screen "2#电梯状态画面" 800x600
   TextField "文本域_1" at 385,17 size 267x27; Text '-- 2#电梯状态总览'
   TextField "文本域_3" at 77,12 size 300x31; Text '电 梯 监 控 系 统'
   Button "按钮_7" at 555,516 size 117x66; TextOff '电梯状态总览'
      on Click: ActivateScreen("电梯状态总览画面", 0)
   Button "按钮_8" at 677,516 size 106x66; TextOff '退出系统'
      on Click: StopRuntime(0)
   Rectangle "矩形_237" at 73,319 size 44x21
      Appearance <- "输出_2号梯5层按钮指示灯"
   Rectangle "矩形_238" at 73,297 size 44x21
      Appearance <- "输出_2号梯6层按钮指示灯"
   Rectangle "矩形_239" at 73,275 size 44x21
      Appearance <- "输出_2号梯7层按钮指示灯"
   Rectangle "矩形_240" at 73,253 size 44x21
      Appearance <- "输出_2号梯8层按钮指示灯"
   Rectangle "矩形_241" at 73,231 size 44x21
      Appearance <- "输出_2号梯9层按钮指示灯"
   Rectangle "矩形_242" at 73,209 size 44x21
      Appearance <- "输出_2号梯10层按钮指示灯"
   Circle "圆_1" at 162,212 size 14x14
      Appearance <- "输出_10层下行呼梯按钮指示灯"
   Circle "圆_2" at 149,234 size 14x14
      Appearance <- "输出_9层上行呼梯按钮指示灯"
   Circle "圆_3" at 174,234 size 14x14
      Appearance <- "输出_9层下行呼梯按钮指示灯"
   Circle "圆_4" at 149,256 size 14x14
      Appearance <- "输出_8层上行呼梯按钮指示灯"
   Circle "圆_5" at 174,256 size 14x14
      Appearance <- "输出_8层下行呼梯按钮指示灯"
   Circle "圆_6" at 149,278 size 14x14
      Appearance <- "输出_7层上行呼梯按钮指示灯"
   Circle "圆_7" at 174,278 size 14x14
      Appearance <- "输出_7层下行呼梯按钮指示灯"
   Circle "圆_8" at 149,299 size 14x14
      Appearance <- "输出_6层上行呼梯按钮指示灯"
   Circle "圆_9" at 174,299 size 14x14
      Appearance <- "输出_6层下行呼梯按钮指示灯"
   Circle "圆_10" at 149,321 size 14x14
      Appearance <- "输出_5层上行呼梯按钮指示灯"
   Circle "圆_11" at 174,321 size 14x14
      Appearance <- "输出_5层下行呼梯按钮指示灯"
   Circle "圆_12" at 149,343 size 14x14
      Appearance <- "输出_4层上行呼梯按钮指示灯"
   Circle "圆_13" at 174,343 size 14x14
      Appearance <- "输出_4层下行呼梯按钮指示灯"
   Circle "圆_14" at 149,365 size 14x14
      Appearance <- "输出_3层上行呼梯按钮指示灯"
   Circle "圆_15" at 174,365 size 14x14
      Appearance <- "输出_3层下行呼梯按钮指示灯"
   Circle "圆_16" at 149,389 size 14x14
      Appearance <- "输出_2层上行呼梯按钮指示灯"
   Circle "圆_17" at 174,389 size 14x14
      Appearance <- "输出_2层下行呼梯按钮指示灯"
   Circle "圆_18" at 162,411 size 14x14
      Appearance <- "输出_1层上行呼梯按钮指示灯"
   TextField "文本域_41" at 75,440 size 45x23; Text '内呼'
   TextField "文本域_42" at 151,441 size 48x24; Text '外呼'
   Rectangle "矩形_233" at 73,407 size 44x21
      Appearance <- "输出_2号梯1层按钮指示灯"
   Rectangle "矩形_234" at 73,385 size 44x21
      Appearance <- "输出_2号梯2层按钮指示灯"
   Button "FB_Empty_Rectangular_1" at 80,409 size 29x18; TextOff 'Text'; PictureOff "FB_Empty_Rectangular_Released_256c"; PictureOn "FB_Empty_Rectangular_Pressed_256c"
      on Release: ResetBit("输入_2号梯轿内选层按钮1")
      on Press: SetBit("输入_2号梯轿内选层按钮1")
   Button "FB_Empty_Rectangular_2" at 81,387 size 29x18; TextOff 'Text'; PictureOff "FB_Empty_Rectangular_Released_256c"; PictureOn "FB_Empty_Rectangular_Pressed_256c"
      on Release: ResetBit("输入_2号梯轿内选层按钮2")
      on Press: SetBit("输入_2号梯轿内选层按钮2")
   Rectangle "矩形_235" at 73,363 size 44x21
      Appearance <- "输出_2号梯3层按钮指示灯"
   Button "FB_Empty_Rectangular_3" at 81,365 size 29x18; TextOff 'Text'; PictureOff "FB_Empty_Rectangular_Released_256c"; PictureOn "FB_Empty_Rectangular_Pressed_256c"
      on Release: ResetBit("输入_2号梯轿内选层按钮3")
      on Press: SetBit("输入_2号梯轿内选层按钮3")
   Rectangle "矩形_236" at 73,341 size 44x21
      Appearance <- "输出_2号梯4层按钮指示灯"
   Button "FB_Empty_Rectangular_4" at 81,343 size 29x18; TextOff 'Text'; PictureOff "FB_Empty_Rectangular_Released_256c"; PictureOn "FB_Empty_Rectangular_Pressed_256c"
      on Release: ResetBit("输入_2号梯轿内选层按钮4")
      on Press: SetBit("输入_2号梯轿内选层按钮4")
   Button "FB_Empty_Rectangular_5" at 81,321 size 29x18; TextOff 'Text'; PictureOff "FB_Empty_Rectangular_Released_256c"; PictureOn "FB_Empty_Rectangular_Pressed_256c"
      on Release: ResetBit("输入_2号梯轿内选层按钮5")
      on Press: SetBit("输入_2号梯轿内选层按钮5")
   Button "FB_Empty_Rectangular_6" at 81,299 size 29x18; TextOff 'Text'; PictureOff "FB_Empty_Rectangular_Released_256c"; PictureOn "FB_Empty_Rectangular_Pressed_256c"
      on Release: ResetBit("输入_2号梯轿内选层按钮6")
      on Press: SetBit("输入_2号梯轿内选层按钮6")
   Button "FB_Empty_Rectangular_7" at 81,277 size 29x18; TextOff 'Text'; PictureOff "FB_Empty_Rectangular_Released_256c"; PictureOn "FB_Empty_Rectangular_Pressed_256c"
      on Release: ResetBit("输入_2号梯轿内选层按钮7")
      on Press: SetBit("输入_2号梯轿内选层按钮7")
   Button "FB_Empty_Rectangular_8" at 81,255 size 29x18; TextOff 'Text'; PictureOff "FB_Empty_Rectangular_Released_256c"; PictureOn "FB_Empty_Rectangular_Pressed_256c"
      on Release: ResetBit("输入_2号梯轿内选层按钮8")
      on Press: SetBit("输入_2号梯轿内选层按钮8")
   Button "FB_Empty_Rectangular_9" at 81,233 size 29x18; TextOff 'Text'; PictureOff "FB_Empty_Rectangular_Released_256c"; PictureOn "FB_Empty_Rectangular_Pressed_256c"
      on Release: ResetBit("输入_2号梯轿内选层按钮9")
      on Press: SetBit("输入_2号梯轿内选层按钮9")
   Button "FB_Empty_Rectangular_10" at 81,211 size 29x18; TextOff 'Text'; PictureOff "FB_Empty_Rectangular_Released_256c"; PictureOn "FB_Empty_Rectangular_Pressed_256c"
      on Release: ResetBit("输入_2号梯轿内选层按钮10")
      on Press: SetBit("输入_2号梯轿内选层按钮10")
   TextField "文本域_14" at 88,409 size 14x19; Text '1'
   TextField "文本域_15" at 88,386 size 14x19; Text '2'
   TextField "文本域_16" at 88,363 size 14x19; Text '3'
   TextField "文本域_17" at 88,342 size 14x19; Text '4'
   TextField "文本域_18" at 88,320 size 14x19; Text '5'
   TextField "文本域_19" at 88,298 size 14x19; Text '6'
   TextField "文本域_20" at 88,276 size 14x19; Text '7'
   TextField "文本域_21" at 88,254 size 14x19; Text '8'
   TextField "文本域_22" at 88,232 size 14x19; Text '9'
   TextField "文本域_40" at 84,210 size 23x19; Text '10'
   Circle "圆_56" at 464,117 size 24x24
      Appearance <- "输出_2号梯满载指示"
   Circle "圆_57" at 574,117 size 24x24
      Appearance <- "输出_2号梯故障指示"
   Circle "圆_58" at 464,164 size 24x24
      Appearance <- "输出_2号梯照明指示"
   Circle "圆_59" at 349,120 size 24x24
      Appearance <- "输出_2号梯满载指示"
   Circle "圆_60" at 575,166 size 24x24
      Appearance <- "输出_2号梯风扇指示"
   TextField "文本域_47" at 383,122 size 37x19; Text '超重'
   TextField "文本域_48" at 498,120 size 61x23; Text '满载'
   TextField "文本域_49" at 608,118 size 50x28; Text '故障'
   TextField "文本域_50" at 502,167 size 54x26; Text '照明'
   TextField "文本域_51" at 609,162 size 58x28; Text '风扇'
   Circle "圆_73" at 215,119 size 24x24
      Appearance <- "输入_自动运行信号"
   TextField "文本域_68" at 246,120 size 87x20; Text '自动运行'
   Group "Group" at 310,468 size 40x20; PictureOn "FB_Left_Square_Pressed_256c"; PictureOff "FB_Left_Square_Released_256c"
   Group "Group_1" at 356,468 size 40x20; PictureOn "FB_Left_Square_Pressed_256c"; PictureOff "FB_Left_Square_Released_256c"
   TextField "文本域_69" at 245,167 size 127x20; Text '电梯准备就绪'
   Circle "圆_83" at 624,288 size 16x16
      Appearance <- "输出_2号梯开门继电器"
   Circle "圆_86" at 624,303 size 16x16
      Appearance <- "输出_2号梯关门继电器"
   Circle "圆_89" at 472,373 size 16x16
      Appearance <- "输入_2号梯开门到位"
   Circle "圆_92" at 472,389 size 16x16
      Appearance <- "输入_2号梯关门到位"
   Circle "圆_129" at 624,238 size 16x16
      Appearance <- "输出_2号梯电机启动信号"
   Circle "圆_132" at 624,253 size 16x16
      Appearance <- "输出_2号梯上行接触器"
   Circle "圆_135" at 624,268 size 16x16
      Appearance <- "输出_2号梯下行接触器"
   Circle "圆_19" at 215,163 size 24x24
      Appearance <- "输出_准备就绪信号"
   Circle "圆_95" at 624,358 size 16x16
      Appearance <- "输出_2号梯1级减速制动"
   Circle "圆_98" at 624,373 size 16x16
      Appearance <- "输出_2号梯2级减速制动"
   Circle "圆_101" at 624,388 size 16x16
      Appearance <- "输出_2号梯3级减速制动"
   Circle "圆_104" at 624,327 size 16x16
      Appearance <- "输出_2号梯低速接触器"
   Circle "圆_107" at 624,342 size 16x16
      Appearance <- "输出_2号梯高速接触器"
   Circle "圆_120" at 317,389 size 16x16
      Appearance <- "输入_2号梯轿厢门锁信号"
   Circle "圆_123" at 317,234 size 16x16
      Appearance <- "输入_2号梯10楼层门锁信号"
   Circle "圆_126" at 317,249 size 16x16
      Appearance <- "输入_2号梯9楼层门锁信号"
   Circle "圆_138" at 317,264 size 16x16
      Appearance <- "输入_2号梯8楼层门锁信号"
   Circle "圆_141" at 317,279 size 16x16
      Appearance <- "输入_2号梯7楼层门锁信号"
   Circle "圆_144" at 317,295 size 16x16
      Appearance <- "输入_2号梯6楼层门锁信号"
   Circle "圆_147" at 317,310 size 16x16
      Appearance <- "输入_2号梯5楼层门锁信号"
   Circle "圆_150" at 317,326 size 16x16
      Appearance <- "输入_2号梯4楼层门锁信号"
   Circle "圆_153" at 317,342 size 16x16
      Appearance <- "输入_2号梯3楼层门锁信号"
   Circle "圆_156" at 317,357 size 16x16
      Appearance <- "输入_2号梯2楼层门锁信号"
   Circle "圆_159" at 317,373 size 16x16
      Appearance <- "输入_2号梯1楼层门锁信号"
   Circle "圆_162" at 472,234 size 16x16
      Appearance <- "输入_2号梯上端站第2限位"
   Circle "圆_165" at 472,249 size 16x16
      Appearance <- "输入_2号梯上端站第1限位"
   Circle "圆_168" at 472,264 size 16x16
      Appearance <- "输入_2号梯上平层信号"
   Circle "圆_171" at 472,279 size 16x16
      Appearance <- "输入_2号梯下平层信号"
   Circle "圆_174" at 472,294 size 16x16
      Appearance <- "输入_2号梯下端站第2限位"
   Circle "圆_177" at 472,309 size 16x16
      Appearance <- "输入_2号梯下端站第1限位"
   Circle "圆_183" at 472,333 size 16x16
      Appearance <- "输入_2号梯检修信号"
   Circle "圆_186" at 472,348 size 16x16
      Appearance <- "输入_2号梯光幕信号"
   Rectangle "矩形_193" at 165,134 size 4x18
      Appearance <- "输出_2号梯LEDi"
   Rectangle "矩形_194" at 165,156 size 4x18
      Appearance <- "输出_2号梯LEDj"
   Rectangle "矩形_195" at 178,132 size 18x4
      Appearance <- "输出_2号梯LEDa"
   Rectangle "矩形_196" at 175,136 size 4x18
      Appearance <- "输出_2号梯LEDf"
   Rectangle "矩形_197" at 178,153 size 18x4
      Appearance <- "输出_2号梯LEDg"
   Rectangle "矩形_198" at 175,157 size 4x18
      Appearance <- "输出_2号梯LEDe"
   Rectangle "矩形_199" at 178,175 size 18x4
      Appearance <- "输出_2号梯LEDd"
   Rectangle "矩形_200" at 195,135 size 4x18
      Appearance <- "输出_2号梯LEDb"
   Rectangle "矩形_201" at 195,157 size 4x18
      Appearance <- "输出_2号梯LEDc"
   Rectangle "矩形_72" at 91,122 size 6x34
      Appearance <- "输出_2号梯上行指示"
   Polygon "多边形_5" at 79,118 size 15x17
      Appearance <- "输出_2号梯上行指示"
   Polygon "多边形_6" at 94,118 size 14x17
      Appearance <- "输出_2号梯上行指示"
   Rectangle "矩形_73" at 91,157 size 6x34
      Appearance <- "输出_2号梯下行指示"
   Polygon "多边形_1" at 77,179 size 17x15
      Appearance <- "输出_2号梯下行指示"
   Polygon "多边形_2" at 94,179 size 17x15
      Appearance <- "输出_2号梯下行指示"
   TextField "文本域_77" at 223,251 size 81x15; Text '9层门锁信号'
   TextField "文本域_78" at 223,266 size 81x15; Text '8层门锁信号'
   TextField "文本域_79" at 223,282 size 81x15; Text '7层门锁信号'
   TextField "文本域_80" at 223,298 size 81x15; Text '6层门锁信号'
   TextField "文本域_81" at 223,314 size 81x15; Text '5层门锁信号'
   TextField "文本域_83" at 223,329 size 81x15; Text '4层门锁信号'
   TextField "文本域_84" at 223,344 size 81x15; Text '3层门锁信号'
   TextField "文本域_85" at 223,360 size 81x15; Text '2层门锁信号'
   TextField "文本域_86" at 222,375 size 82x15; Text '1层门锁信号'
   TextField "文本域_87" at 223,391 size 81x15; Text '轿厢门锁信号'
   TextField "文本域_23" at 382,336 size 72x15; Text '检修开关'
   TextField "文本域_24" at 384,352 size 70x15; Text '光幕信号'
   TextField "文本域_82" at 351,237 size 103x15; Text '上端站第二限位'
   TextField "文本域_88" at 350,255 size 104x15; Text '上端站第一限位'
   TextField "文本域_89" at 372,270 size 82x15; Text '上平层信号'
   TextField "文本域_90" at 372,285 size 82x15; Text '下平层信号'
   TextField "文本域_91" at 350,299 size 104x15; Text '下端站第二限位'
   TextField "文本域_92" at 350,315 size 104x15; Text '下端站第一限位'
   TextField "文本域_13" at 362,372 size 93x15; Text '开门到位信号'
   TextField "文本域_25" at 362,388 size 93x15; Text '关门到位信号'
   TextField "文本域_97" at 525,289 size 92x15; Text '开门继电器'
   TextField "文本域_98" at 525,305 size 92x15; Text '关门继电器'
   TextField "文本域_104" at 525,270 size 92x15; Text '下行接触器'
   TextField "文本域_105" at 514,238 size 103x15; Text '电机启动信号'
   TextField "文本域_106" at 525,254 size 92x15; Text '上行接触器'
   TextField "文本域_99" at 504,374 size 114x15; Text '二级制动接触器'
   TextField "文本域_100" at 504,390 size 114x15; Text '三级制动接触器'
   TextField "文本域_101" at 504,357 size 114x15; Text '一级制动接触器'
   TextField "文本域_102" at 504,325 size 114x15; Text '低速运行接触器'
   TextField "文本域_103" at 504,341 size 114x15; Text '高速运行接触器'
   TextField "文本域_76" at 217,236 size 91x15; Text '10层门锁信号'
   Clock "时钟_1" at 664,57 size 101x57
   DateTimeField "日期/时间域_1" at 491,71 size 184x28
   TextField "文本域_26" at 278,421 size 142x19; Text '1号电梯开关门状态'
   Button "FB_Left_Square" at 310,468 size 20x20; TextOff 'Text'; PictureOff "FB_Left_Square_Released_256c"; PictureOn "FB_Left_Square_Pressed_256c"
      on Click: SetBit("输入_1号梯轿内开门按钮")
      Appearance <- "输入_2号梯轿内关门按钮"
   Button "FB_Right_Square" at 330,468 size 20x20; TextOff 'Text'; PictureOff "FB_Right_Square_Released_256c_2"; PictureOn "FB_Right_Square_Pressed_256c"
      on Click: SetBit("输入_1号梯轿内开门按钮")
      Appearance <- "输入_1号梯轿内开门按钮"
   Button "FB_Left_Square_1" at 376,468 size 20x20; TextOff 'Text'; PictureOff "FB_Left_Square_Released_256c"; PictureOn "FB_Left_Square_Pressed_256c"
      on Click: SetBit("输入_1号梯轿内关门按钮")
      Appearance <- "输入_2号梯轿内关门按钮"
   Button "FB_Right_Square_1" at 356,468 size 20x20; TextOff 'Text'; PictureOff "FB_Right_Square_Released_256c_2"; PictureOn "FB_Right_Square_Pressed_256c"
      on Click: SetBit("输入_1号梯轿内关门按钮")
      Appearance <- "输入_1号梯轿内关门按钮"

screen "3#电梯状态画面" 800x600
   TextField "文本域_1" at 385,17 size 263x27; Text '-- 3#电梯状态总览'
   TextField "文本域_3" at 82,12 size 295x31; Text '电 梯 监 控 系 统'
   Button "按钮_7" at 550,517 size 115x66; TextOff '电梯状态总览'
      on Click: ActivateScreen("电梯状态总览画面", 0)
   Button "按钮_8" at 671,517 size 106x66; TextOff '退出系统'
      on Click: StopRuntime(0)
   Group "Group" at 272,465 size 40x20; PictureOn "FB_Left_Square_Pressed_256c"; PictureOff "FB_Left_Square_Released_256c"
   Group "Group_1" at 324,465 size 40x20; PictureOn "FB_Left_Square_Pressed_256c"; PictureOff "FB_Left_Square_Released_256c"
   Rectangle "矩形_237" at 75,319 size 44x21
      Appearance <- "输出_3号梯5层按钮指示灯"
   Rectangle "矩形_238" at 75,297 size 44x21
      Appearance <- "输出_3号梯6层按钮指示灯"
   Rectangle "矩形_239" at 75,275 size 44x21
      Appearance <- "输出_3号梯7层按钮指示灯"
   Rectangle "矩形_240" at 75,253 size 44x21
      Appearance <- "输出_3号梯8层按钮指示灯"
   Rectangle "矩形_241" at 75,231 size 44x21
      Appearance <- "输出_3号梯9层按钮指示灯"
   Rectangle "矩形_242" at 75,209 size 44x21
      Appearance <- "输出_3号梯10层按钮指示灯"
   Circle "圆_1" at 164,212 size 14x14
      Appearance <- "输出_10层下行呼梯按钮指示灯"
   Circle "圆_2" at 151,232 size 14x14
      Appearance <- "输出_9层上行呼梯按钮指示灯"
   Circle "圆_3" at 176,232 size 14x14
      Appearance <- "输出_9层下行呼梯按钮指示灯"
   Circle "圆_4" at 151,254 size 14x14
      Appearance <- "输出_8层上行呼梯按钮指示灯"
   Circle "圆_5" at 176,254 size 14x14
      Appearance <- "输出_8层下行呼梯按钮指示灯"
   Circle "圆_6" at 151,277 size 14x14
      Appearance <- "输出_7层上行呼梯按钮指示灯"
   Circle "圆_7" at 176,277 size 14x14
      Appearance <- "输出_7层下行呼梯按钮指示灯"
   Circle "圆_8" at 151,299 size 14x14
      Appearance <- "输出_6层上行呼梯按钮指示灯"
   Circle "圆_9" at 176,299 size 14x14
      Appearance <- "输出_6层下行呼梯按钮指示灯"
   Circle "圆_10" at 151,322 size 14x14
      Appearance <- "输出_5层上行呼梯按钮指示灯"
   Circle "圆_11" at 176,322 size 14x14
      Appearance <- "输出_5层下行呼梯按钮指示灯"
   Circle "圆_12" at 151,345 size 14x14
      Appearance <- "输出_4层上行呼梯按钮指示灯"
   Circle "圆_13" at 176,345 size 14x14
      Appearance <- "输出_4层下行呼梯按钮指示灯"
   Circle "圆_14" at 151,367 size 14x14
      Appearance <- "输出_3层上行呼梯按钮指示灯"
   Circle "圆_15" at 176,367 size 14x14
      Appearance <- "输出_3层下行呼梯按钮指示灯"
   Circle "圆_16" at 151,389 size 14x14
      Appearance <- "输出_2层上行呼梯按钮指示灯"
   Circle "圆_17" at 176,389 size 14x14
      Appearance <- "输出_2层下行呼梯按钮指示灯"
   Circle "圆_18" at 163,411 size 14x14
      Appearance <- "输出_1层上行呼梯按钮指示灯"
   TextField "文本域_41" at 77,440 size 45x23; Text '内呼'
   TextField "文本域_42" at 152,440 size 45x23; Text '外呼'
   Rectangle "矩形_233" at 75,407 size 44x21
      Appearance <- "输出_3号梯1层按钮指示灯"
   Rectangle "矩形_234" at 75,385 size 44x21
      Appearance <- "输出_3号梯2层按钮指示灯"
   Button "FB_Empty_Rectangular_1" at 82,410 size 29x18; TextOff 'Text'; PictureOff "FB_Empty_Rectangular_Released_256c"; PictureOn "FB_Empty_Rectangular_Pressed_256c"
      on Release: ResetBit("输入_3号梯轿内选层按钮1")
      on Press: SetBit("输入_3号梯轿内选层按钮1")
      Appearance <- "输出_1号梯1层按钮指示灯"
   Button "FB_Empty_Rectangular_2" at 83,387 size 29x18; TextOff 'Text'; PictureOff "FB_Empty_Rectangular_Released_256c"; PictureOn "FB_Empty_Rectangular_Pressed_256c"
      on Release: ResetBit("输入_3号梯轿内选层按钮2")
      on Press: SetBit("输入_3号梯轿内选层按钮2")
   Rectangle "矩形_235" at 75,363 size 44x21
      Appearance <- "输出_3号梯3层按钮指示灯"
   Button "FB_Empty_Rectangular_3" at 83,365 size 29x18; TextOff 'Text'; PictureOff "FB_Empty_Rectangular_Released_256c"; PictureOn "FB_Empty_Rectangular_Pressed_256c"
      on Release: ResetBit("输入_3号梯轿内选层按钮3")
      on Press: SetBit("输入_3号梯轿内选层按钮3")
   Rectangle "矩形_236" at 75,341 size 44x21
      Appearance <- "输出_3号梯4层按钮指示灯"
   Button "FB_Empty_Rectangular_4" at 83,343 size 29x18; TextOff 'Text'; PictureOff "FB_Empty_Rectangular_Released_256c"; PictureOn "FB_Empty_Rectangular_Pressed_256c"
      on Release: ResetBit("输入_3号梯轿内选层按钮4")
      on Press: SetBit("输入_3号梯轿内选层按钮4")
   Button "FB_Empty_Rectangular_5" at 83,321 size 29x18; TextOff 'Text'; PictureOff "FB_Empty_Rectangular_Released_256c"; PictureOn "FB_Empty_Rectangular_Pressed_256c"
      on Release: ResetBit("输入_3号梯轿内选层按钮5")
      on Press: SetBit("输入_3号梯轿内选层按钮5")
   Button "FB_Empty_Rectangular_6" at 83,299 size 29x18; TextOff 'Text'; PictureOff "FB_Empty_Rectangular_Released_256c"; PictureOn "FB_Empty_Rectangular_Pressed_256c"
      on Release: ResetBit("输入_3号梯轿内选层按钮6")
      on Press: SetBit("输入_3号梯轿内选层按钮6")
   Button "FB_Empty_Rectangular_7" at 83,277 size 29x18; TextOff 'Text'; PictureOff "FB_Empty_Rectangular_Released_256c"; PictureOn "FB_Empty_Rectangular_Pressed_256c"
      on Release: ResetBit("输入_3号梯轿内选层按钮7")
      on Press: SetBit("输入_3号梯轿内选层按钮7")
   Button "FB_Empty_Rectangular_8" at 83,255 size 29x18; TextOff 'Text'; PictureOff "FB_Empty_Rectangular_Released_256c"; PictureOn "FB_Empty_Rectangular_Pressed_256c"
      on Release: ResetBit("输入_3号梯轿内选层按钮8")
      on Press: SetBit("输入_3号梯轿内选层按钮8")
   Button "FB_Empty_Rectangular_9" at 83,233 size 29x18; TextOff 'Text'; PictureOff "FB_Empty_Rectangular_Released_256c"; PictureOn "FB_Empty_Rectangular_Pressed_256c"
      on Release: ResetBit("输入_3号梯轿内选层按钮9")
      on Press: SetBit("输入_3号梯轿内选层按钮9")
   Button "FB_Empty_Rectangular_10" at 83,211 size 29x18; TextOff 'Text'; PictureOff "FB_Empty_Rectangular_Released_256c"; PictureOn "FB_Empty_Rectangular_Pressed_256c"
      on Release: ResetBit("输入_3号梯轿内选层按钮10")
      on Press: SetBit("输入_3号梯轿内选层按钮10")
   TextField "文本域_14" at 90,409 size 14x19; Text '1'
   TextField "文本域_15" at 90,386 size 14x19; Text '2'
   TextField "文本域_16" at 90,363 size 14x19; Text '3'
   TextField "文本域_17" at 90,342 size 14x19; Text '4'
   TextField "文本域_18" at 90,320 size 14x19; Text '5'
   TextField "文本域_19" at 90,298 size 14x19; Text '6'
   TextField "文本域_20" at 90,276 size 14x19; Text '7'
   TextField "文本域_21" at 90,254 size 14x19; Text '8'
   TextField "文本域_22" at 90,232 size 14x19; Text '9'
   TextField "文本域_40" at 86,210 size 23x19; Text '10'
   Circle "圆_56" at 476,117 size 24x24
      Appearance <- "输出_3号梯满载指示"
   Circle "圆_57" at 586,117 size 24x24
      Appearance <- "输出_3号梯故障指示"
   Circle "圆_58" at 476,166 size 24x24
      Appearance <- "输出_3号梯照明指示"
   Circle "圆_59" at 372,119 size 24x24
      Appearance <- "输出_3号梯满载指示"
   Circle "圆_60" at 587,168 size 24x24
      Appearance <- "输出_3号梯风扇指示"
   TextField "文本域_47" at 403,119 size 45x23; Text '超重'
   TextField "文本域_48" at 510,120 size 45x23; Text '满载'
   TextField "文本域_49" at 622,119 size 45x23; Text '故障'
   TextField "文本域_50" at 514,169 size 45x23; Text '照明'
   TextField "文本域_51" at 624,168 size 45x23; Text '风扇'
   Circle "圆_73" at 227,119 size 24x24
      Appearance <- "输入_自动运行信号"
   TextField "文本域_68" at 258,120 size 73x20; Text '自动运行'
   TextField "文本域_69" at 257,167 size 107x20; Text '电梯准备就绪'
   Circle "圆_83" at 625,280 size 16x16
      Appearance <- "输出_3号梯开门继电器"
   Circle "圆_86" at 625,295 size 16x16
      Appearance <- "输出_3号梯关门继电器"
   Circle "圆_89" at 477,363 size 16x16
      Appearance <- "输入_3号梯开门到位"
   Circle "圆_92" at 477,379 size 16x16
      Appearance <- "输入_3号梯关门到位"
   Circle "圆_129" at 624,229 size 16x16
      Appearance <- "输出_3号梯电机启动信号"
   Circle "圆_132" at 624,244 size 16x16
      Appearance <- "输出_3号梯上行接触器"
   Circle "圆_135" at 624,259 size 16x16
      Appearance <- "输出_3号梯下行接触器"
   Circle "圆_19" at 227,163 size 24x24
      Appearance <- "输出_准备就绪信号"
   Circle "圆_95" at 625,352 size 16x16
      Appearance <- "输出_3号梯1级减速制动"
   Circle "圆_98" at 625,367 size 16x16
      Appearance <- "输出_3号梯2级减速制动"
   Circle "圆_101" at 625,382 size 16x16
      Appearance <- "输出_3号梯3级减速制动"
   Circle "圆_104" at 625,321 size 16x16
      Appearance <- "输出_3号梯低速接触器"
   Circle "圆_107" at 625,336 size 16x16
      Appearance <- "输出_3号梯高速接触器"
   Circle "圆_120" at 324,378 size 16x16
      Appearance <- "输入_3号梯轿厢门锁信号"
   Circle "圆_123" at 324,228 size 16x16
      Appearance <- "输入_3号梯10楼层门锁信号"
   Circle "圆_126" at 324,243 size 16x16
      Appearance <- "输入_3号梯9楼层门锁信号"
   Circle "圆_138" at 324,258 size 16x16
      Appearance <- "输入_3号梯8楼层门锁信号"
   Circle "圆_141" at 324,273 size 16x16
      Appearance <- "输入_3号梯7楼层门锁信号"
   Circle "圆_144" at 324,288 size 16x16
      Appearance <- "输入_3号梯6楼层门锁信号"
   Circle "圆_147" at 324,303 size 16x16
      Appearance <- "输入_3号梯5楼层门锁信号"
   Circle "圆_150" at 324,318 size 16x16
      Appearance <- "输入_3号梯4楼层门锁信号"
   Circle "圆_153" at 324,333 size 16x16
      Appearance <- "输入_3号梯3楼层门锁信号"
   Circle "圆_156" at 324,348 size 16x16
      Appearance <- "输入_3号梯2楼层门锁信号"
   Circle "圆_159" at 324,363 size 16x16
      Appearance <- "输入_3号梯1楼层门锁信号"
   Circle "圆_162" at 476,228 size 16x16
      Appearance <- "输入_3号梯上端站第2限位"
   Circle "圆_165" at 476,243 size 16x16
      Appearance <- "输入_3号梯上端站第1限位"
   Circle "圆_168" at 476,258 size 16x16
      Appearance <- "输入_3号梯上平层信号"
   Circle "圆_171" at 476,273 size 16x16
      Appearance <- "输入_3号梯下平层信号"
   Circle "圆_174" at 476,288 size 16x16
      Appearance <- "输入_3号梯下端站第2限位"
   Circle "圆_177" at 476,303 size 16x16
      Appearance <- "输入_3号梯下端站第1限位"
   Circle "圆_183" at 476,327 size 16x16
      Appearance <- "输入_3号梯检修信号"
   Circle "圆_186" at 476,342 size 16x16
      Appearance <- "输入_3号梯光幕信号"
   Rectangle "矩形_193" at 167,134 size 4x18
      Appearance <- "输出_3号梯LEDi"
   Rectangle "矩形_194" at 167,156 size 4x18
      Appearance <- "输出_3号梯LEDj"
   Rectangle "矩形_195" at 180,132 size 18x4
      Appearance <- "输出_3号梯LEDa"
   Rectangle "矩形_196" at 177,136 size 4x18
      Appearance <- "输出_3号梯LEDf"
   Rectangle "矩形_197" at 180,153 size 18x4
      Appearance <- "输出_3号梯LEDg"
   Rectangle "矩形_198" at 177,157 size 4x18
      Appearance <- "输出_3号梯LEDe"
   Rectangle "矩形_199" at 180,175 size 18x4
      Appearance <- "输出_3号梯LEDd"
   Rectangle "矩形_200" at 197,135 size 4x18
      Appearance <- "输出_3号梯LEDb"
   Rectangle "矩形_201" at 197,157 size 4x18
      Appearance <- "输出_3号梯LEDc"
   Rectangle "矩形_72" at 93,122 size 6x34
      Appearance <- "输出_3号梯上行指示"
   Polygon "多边形_5" at 81,118 size 15x17
      Appearance <- "输出_3号梯上行指示"
   Polygon "多边形_6" at 96,118 size 14x17
      Appearance <- "输出_3号梯上行指示"
   Rectangle "矩形_73" at 93,157 size 6x34
      Appearance <- "输出_3号梯下行指示"
   Polygon "多边形_1" at 79,179 size 17x15
      Appearance <- "输出_3号梯下行指示"
   Polygon "多边形_2" at 96,179 size 17x15
      Appearance <- "输出_3号梯下行指示"
   TextField "文本域_23" at 388,326 size 72x15; Text '检修开关'
   TextField "文本域_24" at 390,342 size 70x15; Text '光幕信号'
   TextField "文本域_82" at 357,229 size 103x15; Text '上端站第二限位'
   TextField "文本域_88" at 356,245 size 104x15; Text '上端站第一限位'
   TextField "文本域_89" at 378,260 size 82x15; Text '上平层信号'
   TextField "文本域_90" at 378,275 size 82x15; Text '下平层信号'
   TextField "文本域_91" at 356,291 size 104x15; Text '下端站第二限位'
   TextField "文本域_92" at 356,307 size 104x15; Text '下端站第一限位'
   TextField "文本域_13" at 368,364 size 93x15; Text '开门到位信号'
   TextField "文本域_25" at 368,380 size 93x15; Text '关门到位信号'
   TextField "文本域_97" at 528,282 size 92x15; Text '开门继电器'
   TextField "文本域_98" at 528,298 size 92x15; Text '关门继电器'
   TextField "文本域_104" at 528,263 size 92x15; Text '下行接触器'
   TextField "文本域_105" at 517,231 size 103x15; Text '电机启动信号'
   TextField "文本域_106" at 528,247 size 92x15; Text '上行接触器'
   TextField "文本域_99" at 507,367 size 114x15; Text '二级制动接触器'
   TextField "文本域_100" at 507,383 size 114x15; Text '三级制动接触器'
   TextField "文本域_101" at 507,350 size 114x15; Text '一级制动接触器'
   TextField "文本域_102" at 507,318 size 114x15; Text '低速运行接触器'
   TextField "文本域_103" at 507,334 size 114x15; Text '高速运行接触器'
   TextField "文本域_76" at 219,229 size 91x15; Text '10层门锁信号'
   TextField "文本域_77" at 225,245 size 81x15; Text '9层门锁信号'
   TextField "文本域_78" at 225,260 size 81x15; Text '8层门锁信号'
   TextField "文本域_79" at 225,274 size 81x15; Text '7层门锁信号'
   TextField "文本域_80" at 225,289 size 81x15; Text '6层门锁信号'
   TextField "文本域_81" at 225,304 size 81x15; Text '5层门锁信号'
   TextField "文本域_83" at 225,319 size 81x15; Text '4层门锁信号'
   TextField "文本域_84" at 225,335 size 81x15; Text '3层门锁信号'
   TextField "文本域_85" at 225,350 size 81x15; Text '2层门锁信号'
   TextField "文本域_86" at 224,365 size 82x15; Text '1层门锁信号'
   TextField "文本域_87" at 225,380 size 81x15; Text '轿厢门锁信号'
   Clock "时钟_1" at 664,57 size 101x57
   DateTimeField "日期/时间域_1" at 491,71 size 184x28
   TextField "文本域_26" at 243,428 size 142x19; Text '1号电梯开关门状态'
   Button "FB_Left_Square" at 272,465 size 20x20; TextOff 'Text'; PictureOff "FB_Left_Square_Released_256c"; PictureOn "FB_Left_Square_Pressed_256c"
      on Click: SetBit("输入_1号梯轿内开门按钮")
      Appearance <- "输入_3号梯轿内开门按钮"
   Button "FB_Right_Square" at 292,465 size 20x20; TextOff 'Text'; PictureOff "FB_Right_Square_Released_256c_3"; PictureOn "FB_Right_Square_Pressed_256c"
      on Click: SetBit("输入_1号梯轿内开门按钮")
      Appearance <- "输入_1号梯轿内开门按钮"
   Button "FB_Left_Square_1" at 344,465 size 20x20; TextOff 'Text'; PictureOff "FB_Left_Square_Released_256c"; PictureOn "FB_Left_Square_Pressed_256c"
      on Click: SetBit("输入_1号梯轿内关门按钮")
      Appearance <- "输入_3号梯轿内关门按钮"
   Button "FB_Right_Square_1" at 324,465 size 20x20; TextOff 'Text'; PictureOff "FB_Right_Square_Released_256c_3"; PictureOn "FB_Right_Square_Pressed_256c"
      on Click: SetBit("输入_1号梯轿内关门按钮")
      Appearance <- "输入_1号梯轿内关门按钮"

screen "4#电梯状态画面" 800x600
   TextField "文本域_1" at 385,17 size 287x27; Text '-- 4#电梯状态总览'
   TextField "文本域_3" at 71,12 size 306x31; Text '电 梯 监 控 系 统'
   Button "按钮_7" at 538,519 size 118x66; TextOff '电梯状态总览'
      on Click: ActivateScreen("电梯状态总览画面", 0)
   Button "按钮_8" at 664,519 size 106x66; TextOff '退出系统'
      on Click: StopRuntime(0)
   Group "Group" at 303,439 size 40x20; PictureOn "FB_Left_Square_Pressed_256c"; PictureOff "FB_Left_Square_Released_256c"
   Group "Group_1" at 349,439 size 40x20; PictureOn "FB_Left_Square_Pressed_256c"; PictureOff "FB_Left_Square_Released_256c"
   Rectangle "矩形_237" at 75,315 size 44x21
      Appearance <- "输出_4号梯5层按钮指示灯"
   Rectangle "矩形_238" at 75,293 size 44x21
      Appearance <- "输出_4号梯6层按钮指示灯"
   Rectangle "矩形_239" at 75,271 size 44x21
      Appearance <- "输出_4号梯7层按钮指示灯"
   Rectangle "矩形_240" at 75,249 size 44x21
      Appearance <- "输出_4号梯8层按钮指示灯"
   Rectangle "矩形_241" at 75,227 size 44x21
      Appearance <- "输出_4号梯9层按钮指示灯"
   Rectangle "矩形_242" at 75,205 size 44x21
      Appearance <- "输出_4号梯10层按钮指示灯"
   Circle "圆_1" at 162,208 size 14x14
      Appearance <- "输出_10层下行呼梯按钮指示灯"
   Circle "圆_2" at 151,230 size 14x14
      Appearance <- "输出_9层上行呼梯按钮指示灯"
   Circle "圆_3" at 176,230 size 14x14
      Appearance <- "输出_9层下行呼梯按钮指示灯"
   Circle "圆_4" at 151,251 size 14x14
      Appearance <- "输出_8层上行呼梯按钮指示灯"
   Circle "圆_5" at 176,251 size 14x14
      Appearance <- "输出_8层下行呼梯按钮指示灯"
   Circle "圆_6" at 151,273 size 14x14
      Appearance <- "输出_7层上行呼梯按钮指示灯"
   Circle "圆_7" at 176,273 size 14x14
      Appearance <- "输出_7层下行呼梯按钮指示灯"
   Circle "圆_8" at 151,296 size 14x14
      Appearance <- "输出_6层上行呼梯按钮指示灯"
   Circle "圆_9" at 176,296 size 14x14
      Appearance <- "输出_6层下行呼梯按钮指示灯"
   Circle "圆_10" at 151,318 size 14x14
      Appearance <- "输出_5层上行呼梯按钮指示灯"
   Circle "圆_11" at 176,318 size 14x14
      Appearance <- "输出_5层下行呼梯按钮指示灯"
   Circle "圆_12" at 151,341 size 14x14
      Appearance <- "输出_4层上行呼梯按钮指示灯"
   Circle "圆_13" at 176,341 size 14x14
      Appearance <- "输出_4层下行呼梯按钮指示灯"
   Circle "圆_14" at 151,364 size 14x14
      Appearance <- "输出_3层上行呼梯按钮指示灯"
   Circle "圆_15" at 176,364 size 14x14
      Appearance <- "输出_3层下行呼梯按钮指示灯"
   Circle "圆_16" at 151,385 size 14x14
      Appearance <- "输出_2层上行呼梯按钮指示灯"
   Circle "圆_17" at 176,385 size 14x14
      Appearance <- "输出_2层下行呼梯按钮指示灯"
   Circle "圆_18" at 164,407 size 14x14
      Appearance <- "输出_1层上行呼梯按钮指示灯"
   TextField "文本域_41" at 77,436 size 45x23; Text '内呼'
   TextField "文本域_42" at 145,434 size 45x23; Text '外呼'
   Rectangle "矩形_233" at 75,403 size 44x21
      Appearance <- "输出_4号梯1层按钮指示灯"
   Rectangle "矩形_234" at 75,381 size 44x21
      Appearance <- "输出_4号梯2层按钮指示灯"
   Button "FB_Empty_Rectangular_1" at 82,406 size 29x18; TextOff 'Text'; PictureOff "FB_Empty_Rectangular_Released_256c"; PictureOn "FB_Empty_Rectangular_Pressed_256c"
      on Release: ResetBit("输入_1号梯轿内选层按钮1")
      on Press: SetBit("输入_1号梯轿内选层按钮1")
   Button "FB_Empty_Rectangular_2" at 83,383 size 29x18; TextOff 'Text'; PictureOff "FB_Empty_Rectangular_Released_256c"; PictureOn "FB_Empty_Rectangular_Pressed_256c"
      on Release: ResetBit("输入_1号梯轿内选层按钮2")
      on Press: SetBit("输入_1号梯轿内选层按钮2")
   Rectangle "矩形_235" at 75,359 size 44x21
      Appearance <- "输出_4号梯3层按钮指示灯"
   Button "FB_Empty_Rectangular_3" at 83,361 size 29x18; TextOff 'Text'; PictureOff "FB_Empty_Rectangular_Released_256c"; PictureOn "FB_Empty_Rectangular_Pressed_256c"
      on Release: ResetBit("输入_1号梯轿内选层按钮3")
      on Press: SetBit("输入_1号梯轿内选层按钮3")
   Rectangle "矩形_236" at 75,337 size 44x21
      Appearance <- "输出_4号梯4层按钮指示灯"
   Button "FB_Empty_Rectangular_4" at 83,339 size 29x18; TextOff 'Text'; PictureOff "FB_Empty_Rectangular_Released_256c"; PictureOn "FB_Empty_Rectangular_Pressed_256c"
      on Release: ResetBit("输入_1号梯轿内选层按钮4")
      on Press: SetBit("输入_1号梯轿内选层按钮4")
   Button "FB_Empty_Rectangular_5" at 83,317 size 29x18; TextOff 'Text'; PictureOff "FB_Empty_Rectangular_Released_256c"; PictureOn "FB_Empty_Rectangular_Pressed_256c"
      on Release: ResetBit("输入_1号梯轿内选层按钮5")
      on Press: SetBit("输入_1号梯轿内选层按钮5")
   Button "FB_Empty_Rectangular_6" at 83,295 size 29x18; TextOff 'Text'; PictureOff "FB_Empty_Rectangular_Released_256c"; PictureOn "FB_Empty_Rectangular_Pressed_256c"
      on Release: ResetBit("输入_1号梯轿内选层按钮6")
      on Press: SetBit("输入_1号梯轿内选层按钮6")
   Button "FB_Empty_Rectangular_7" at 83,273 size 29x18; TextOff 'Text'; PictureOff "FB_Empty_Rectangular_Released_256c"; PictureOn "FB_Empty_Rectangular_Pressed_256c"
      on Release: ResetBit("输入_1号梯轿内选层按钮7")
      on Press: SetBit("输入_1号梯轿内选层按钮7")
   Button "FB_Empty_Rectangular_8" at 83,251 size 29x18; TextOff 'Text'; PictureOff "FB_Empty_Rectangular_Released_256c"; PictureOn "FB_Empty_Rectangular_Pressed_256c"
      on Release: ResetBit("输入_1号梯轿内选层按钮8")
      on Press: SetBit("输入_1号梯轿内选层按钮8")
   Button "FB_Empty_Rectangular_9" at 83,229 size 29x18; TextOff 'Text'; PictureOff "FB_Empty_Rectangular_Released_256c"; PictureOn "FB_Empty_Rectangular_Pressed_256c"
      on Release: ResetBit("输入_1号梯轿内选层按钮9")
      on Press: SetBit("输入_1号梯轿内选层按钮9")
   Button "FB_Empty_Rectangular_10" at 83,207 size 29x18; TextOff 'Text'; PictureOff "FB_Empty_Rectangular_Released_256c"; PictureOn "FB_Empty_Rectangular_Pressed_256c"
      on Release: ResetBit("输入_1号梯轿内选层按钮10")
      on Press: SetBit("输入_1号梯轿内选层按钮10")
   TextField "文本域_14" at 90,405 size 14x19; Text '1'
   TextField "文本域_15" at 90,382 size 14x19; Text '2'
   TextField "文本域_16" at 90,359 size 14x19; Text '3'
   TextField "文本域_17" at 90,338 size 14x19; Text '4'
   TextField "文本域_18" at 90,316 size 14x19; Text '5'
   TextField "文本域_19" at 90,294 size 14x19; Text '6'
   TextField "文本域_20" at 90,272 size 14x19; Text '7'
   TextField "文本域_21" at 90,250 size 14x19; Text '8'
   TextField "文本域_22" at 90,228 size 14x19; Text '9'
   TextField "文本域_40" at 86,206 size 23x19; Text '10'
   Circle "圆_56" at 470,112 size 24x24
      Appearance <- "输出_4号梯满载指示"
   Circle "圆_57" at 580,112 size 24x24
      Appearance <- "输出_4号梯故障指示"
   Circle "圆_58" at 470,156 size 24x24
      Appearance <- "输出_4号梯照明指示"
   Circle "圆_59" at 368,114 size 24x24
      Appearance <- "输出_4号梯满载指示"
   Circle "圆_60" at 581,158 size 24x24
      Appearance <- "输出_4号梯风扇指示"
   TextField "文本域_47" at 397,114 size 45x23; Text '超重'
   TextField "文本域_48" at 504,115 size 45x23; Text '满载'
   TextField "文本域_49" at 616,114 size 45x23; Text '故障'
   TextField "文本域_50" at 508,159 size 45x23; Text '照明'
   TextField "文本域_51" at 618,159 size 45x23; Text '风扇'
   Circle "圆_73" at 221,114 size 24x24
      Appearance <- "输入_自动运行信号"
   TextField "文本域_68" at 252,115 size 73x20; Text '自动运行'
   TextField "文本域_69" at 254,162 size 107x20; Text '电梯准备就绪'
   Circle "圆_83" at 476,348 size 16x16
      Appearance <- "输出_4号梯开门继电器"
   Circle "圆_86" at 476,363 size 16x16
      Appearance <- "输出_4号梯关门继电器"
   Circle "圆_89" at 626,267 size 16x16
      Appearance <- "输入_4号梯开门到位"
   Circle "圆_92" at 626,283 size 16x16
      Appearance <- "输入_4号梯关门到位"
   Circle "圆_129" at 626,214 size 16x16
      Appearance <- "输出_4号梯电机启动信号"
   Circle "圆_132" at 626,229 size 16x16
      Appearance <- "输出_4号梯上行接触器"
   Circle "圆_135" at 626,244 size 16x16
      Appearance <- "输出_4号梯下行接触器"
   Circle "圆_19" at 221,158 size 24x24
      Appearance <- "输出_准备就绪信号"
   Circle "圆_95" at 627,338 size 16x16
      Appearance <- "输出_4号梯1级减速制动"
   Circle "圆_98" at 627,353 size 16x16
      Appearance <- "输出_4号梯2级减速制动"
   Circle "圆_101" at 627,368 size 16x16
      Appearance <- "输出_4号梯3级减速制动"
   Circle "圆_104" at 627,307 size 16x16
      Appearance <- "输出_4号梯低速接触器"
   Circle "圆_107" at 627,322 size 16x16
      Appearance <- "输出_4号梯高速接触器"
   Circle "圆_120" at 331,366 size 16x16
      Appearance <- "输入_4号梯轿厢门锁信号"
   Circle "圆_123" at 331,214 size 16x16
      Appearance <- "输入_4号梯10楼层门锁信号"
   Circle "圆_126" at 331,229 size 16x16
      Appearance <- "输入_4号梯9楼层门锁信号"
   Circle "圆_138" at 331,244 size 16x16
      Appearance <- "输入_4号梯8楼层门锁信号"
   Circle "圆_141" at 331,259 size 16x16
      Appearance <- "输入_4号梯7楼层门锁信号"
   Circle "圆_144" at 331,274 size 16x16
      Appearance <- "输入_4号梯6楼层门锁信号"
   Circle "圆_147" at 331,289 size 16x16
      Appearance <- "输入_4号梯5楼层门锁信号"
   Circle "圆_150" at 331,304 size 16x16
      Appearance <- "输入_4号梯4楼层门锁信号"
   Circle "圆_153" at 331,319 size 16x16
      Appearance <- "输入_4号梯3楼层门锁信号"
   Circle "圆_156" at 331,334 size 16x16
      Appearance <- "输入_4号梯2楼层门锁信号"
   Circle "圆_159" at 331,350 size 16x16
      Appearance <- "输入_4号梯1楼层门锁信号"
   Circle "圆_162" at 476,212 size 16x16
      Appearance <- "输入_4号梯上端站第2限位"
   Circle "圆_165" at 476,227 size 16x16
      Appearance <- "输入_4号梯上端站第1限位"
   Circle "圆_168" at 476,242 size 16x16
      Appearance <- "输入_4号梯上平层信号"
   Circle "圆_171" at 476,257 size 16x16
      Appearance <- "输入_4号梯下平层信号"
   Circle "圆_174" at 476,272 size 16x16
      Appearance <- "输入_4号梯下端站第2限位"
   Circle "圆_177" at 476,287 size 16x16
      Appearance <- "输入_4号梯下端站第1限位"
   Circle "圆_183" at 476,312 size 16x16
      Appearance <- "输入_4号梯检修信号"
   Circle "圆_186" at 476,327 size 16x16
      Appearance <- "输入_4号梯光幕信号"
   Rectangle "矩形_193" at 167,130 size 4x18
      Appearance <- "输出_4号梯LEDi"
   Rectangle "矩形_194" at 167,152 size 4x18
      Appearance <- "输出_4号梯LEDj"
   Rectangle "矩形_195" at 180,128 size 18x4
      Appearance <- "输出_4号梯LEDa"
   Rectangle "矩形_196" at 177,132 size 4x18
      Appearance <- "输出_4号梯LEDf"
   Rectangle "矩形_197" at 180,149 size 18x4
      Appearance <- "输出_4号梯LEDg"
   Rectangle "矩形_198" at 177,153 size 4x18
      Appearance <- "输出_4号梯LEDe"
   Rectangle "矩形_199" at 180,171 size 18x4
      Appearance <- "输出_4号梯LEDd"
   Rectangle "矩形_200" at 197,131 size 4x18
      Appearance <- "输出_4号梯LEDb"
   Rectangle "矩形_201" at 197,153 size 4x18
      Appearance <- "输出_4号梯LEDc"
   Rectangle "矩形_72" at 93,118 size 6x34
      Appearance <- "输出_4号梯上行指示"
   Polygon "多边形_5" at 81,114 size 15x17
      Appearance <- "输出_4号梯上行指示"
   Polygon "多边形_6" at 96,114 size 14x17
      Appearance <- "输出_4号梯上行指示"
   Rectangle "矩形_73" at 93,153 size 6x34
      Appearance <- "输出_4号梯下行指示"
   Polygon "多边形_1" at 79,175 size 17x15
      Appearance <- "输出_4号梯下行指示"
   Polygon "多边形_2" at 96,175 size 17x15
      Appearance <- "输出_4号梯下行指示"
   TextField "文本域_77" at 225,231 size 81x15; Text '9层门锁信号'
   TextField "文本域_78" at 225,245 size 81x15; Text '8层门锁信号'
   TextField "文本域_79" at 225,260 size 81x15; Text '7层门锁信号'
   TextField "文本域_80" at 225,275 size 81x15; Text '6层门锁信号'
   TextField "文本域_81" at 225,290 size 81x15; Text '5层门锁信号'
   TextField "文本域_83" at 225,306 size 81x15; Text '4层门锁信号'
   TextField "文本域_84" at 225,322 size 81x15; Text '3层门锁信号'
   TextField "文本域_85" at 225,337 size 81x15; Text '2层门锁信号'
   TextField "文本域_86" at 224,354 size 82x15; Text '1层门锁信号'
   TextField "文本域_87" at 220,369 size 86x15; Text '轿厢门锁信号'
   TextField "文本域_23" at 399,312 size 72x15; Text '检修开关'
   TextField "文本域_24" at 401,328 size 70x15; Text '光幕信号'
   TextField "文本域_82" at 368,215 size 103x15; Text '上端站第二限位'
   TextField "文本域_88" at 367,231 size 104x15; Text '上端站第一限位'
   TextField "文本域_89" at 389,246 size 82x15; Text '上平层信号'
   TextField "文本域_90" at 389,261 size 82x15; Text '下平层信号'
   TextField "文本域_91" at 367,275 size 104x15; Text '下端站第二限位'
   TextField "文本域_92" at 367,291 size 104x15; Text '下端站第一限位'
   TextField "文本域_13" at 379,348 size 93x15; Text '开门到位信号'
   TextField "文本域_25" at 379,364 size 93x15; Text '关门到位信号'
   TextField "文本域_97" at 531,267 size 92x15; Text '开门继电器'
   TextField "文本域_98" at 531,283 size 92x15; Text '关门继电器'
   TextField "文本域_104" at 531,248 size 92x15; Text '下行接触器'
   TextField "文本域_105" at 520,216 size 103x15; Text '电机启动信号'
   TextField "文本域_106" at 531,232 size 92x15; Text '上行接触器'
   TextField "文本域_99" at 510,352 size 114x15; Text '二级制动接触器'
   TextField "文本域_100" at 510,368 size 114x15; Text '三级制动接触器'
   TextField "文本域_101" at 510,335 size 114x15; Text '一级制动接触器'
   TextField "文本域_102" at 510,303 size 114x15; Text '低速运行接触器'
   TextField "文本域_103" at 510,319 size 114x15; Text '高速运行接触器'
   TextField "文本域_76" at 219,214 size 91x15; Text '10层门锁信号'
   Clock "时钟_1" at 664,57 size 101x57
   DateTimeField "日期/时间域_1" at 491,71 size 184x28
   TextField "文本域_26" at 269,403 size 142x19; Text '1号电梯开关门状态'
   Button "FB_Left_Square" at 303,439 size 20x20; TextOff 'Text'; PictureOff "FB_Left_Square_Released_256c"; PictureOn "FB_Left_Square_Pressed_256c"
      on Click: SetBit("输入_1号梯轿内开门按钮")
      Appearance <- "输入_4号梯轿内开门按钮"
   Button "FB_Right_Square" at 323,439 size 20x20; TextOff 'Text'; PictureOff "FB_Right_Square_Released_256c_4"; PictureOn "FB_Right_Square_Pressed_256c"
      on Click: SetBit("输入_1号梯轿内开门按钮")
      Appearance <- "输入_1号梯轿内开门按钮"
   Button "FB_Left_Square_1" at 369,439 size 20x20; TextOff 'Text'; PictureOff "FB_Left_Square_Released_256c"; PictureOn "FB_Left_Square_Pressed_256c"
      on Click: SetBit("输入_1号梯轿内关门按钮")
      Appearance <- "输入_4号梯轿内关门按钮"
   Button "FB_Right_Square_1" at 349,439 size 20x20; TextOff 'Text'; PictureOff "FB_Right_Square_Released_256c_4"; PictureOn "FB_Right_Square_Pressed_256c"
      on Click: SetBit("输入_1号梯轿内关门按钮")
      Appearance <- "输入_1号梯轿内关门按钮"

screen "5#电梯状态画面" 800x600
   TextField "文本域_1" at 385,17 size 274x27; Text '-- 5#电梯状态总览'
   TextField "文本域_3" at 76,12 size 301x31; Text '电 梯 监 控 系 统'
   Button "按钮_7" at 547,518 size 121x66; TextOff '电梯状态总览'
      on Click: ActivateScreen("电梯状态总览画面", 0)
   Button "按钮_8" at 675,518 size 106x66; TextOff '退出系统'
      on Click: StopRuntime(0)
   Group "Group" at 284,442 size 40x20; PictureOn "FB_Left_Square_Pressed_256c"; PictureOff "FB_Left_Square_Released_256c"
   Group "Group_1" at 330,442 size 40x20; PictureOn "FB_Left_Square_Pressed_256c"; PictureOff "FB_Left_Square_Released_256c"
   Rectangle "矩形_237" at 75,319 size 44x21
      Appearance <- "输出_5号梯5层按钮指示灯"
   Rectangle "矩形_238" at 75,297 size 44x21
      Appearance <- "输出_5号梯6层按钮指示灯"
   Rectangle "矩形_239" at 75,275 size 44x21
      Appearance <- "输出_5号梯7层按钮指示灯"
   Rectangle "矩形_240" at 75,253 size 44x21
      Appearance <- "输出_5号梯8层按钮指示灯"
   Rectangle "矩形_241" at 75,231 size 44x21
      Appearance <- "输出_5号梯9层按钮指示灯"
   Rectangle "矩形_242" at 75,209 size 44x21
      Appearance <- "输出_5号梯10层按钮指示灯"
   Circle "圆_1" at 163,212 size 14x14
      Appearance <- "输出_10层下行呼梯按钮指示灯"
   Circle "圆_2" at 151,233 size 14x14
      Appearance <- "输出_9层上行呼梯按钮指示灯"
   Circle "圆_3" at 176,233 size 14x14
      Appearance <- "输出_9层下行呼梯按钮指示灯"
   Circle "圆_4" at 151,254 size 14x14
      Appearance <- "输出_8层上行呼梯按钮指示灯"
   Circle "圆_5" at 176,254 size 14x14
      Appearance <- "输出_8层下行呼梯按钮指示灯"
   Circle "圆_6" at 151,277 size 14x14
      Appearance <- "输出_7层上行呼梯按钮指示灯"
   Circle "圆_7" at 176,277 size 14x14
      Appearance <- "输出_7层下行呼梯按钮指示灯"
   Circle "圆_8" at 151,299 size 14x14
      Appearance <- "输出_6层上行呼梯按钮指示灯"
   Circle "圆_9" at 176,299 size 14x14
      Appearance <- "输出_6层下行呼梯按钮指示灯"
   Circle "圆_10" at 151,322 size 14x14
      Appearance <- "输出_5层上行呼梯按钮指示灯"
   Circle "圆_11" at 176,322 size 14x14
      Appearance <- "输出_5层下行呼梯按钮指示灯"
   Circle "圆_12" at 151,345 size 14x14
      Appearance <- "输出_4层上行呼梯按钮指示灯"
   Circle "圆_13" at 176,345 size 14x14
      Appearance <- "输出_4层下行呼梯按钮指示灯"
   Circle "圆_14" at 151,366 size 14x14
      Appearance <- "输出_3层上行呼梯按钮指示灯"
   Circle "圆_15" at 176,366 size 14x14
      Appearance <- "输出_3层下行呼梯按钮指示灯"
   Circle "圆_16" at 151,389 size 14x14
      Appearance <- "输出_2层上行呼梯按钮指示灯"
   Circle "圆_17" at 176,389 size 14x14
      Appearance <- "输出_2层下行呼梯按钮指示灯"
   Circle "圆_18" at 163,411 size 14x14
      Appearance <- "输出_1层上行呼梯按钮指示灯"
   TextField "文本域_41" at 77,440 size 45x23; Text '内呼'
   TextField "文本域_42" at 153,438 size 45x23; Text '外呼'
   Rectangle "矩形_233" at 75,407 size 44x21
      Appearance <- "输出_5号梯1层按钮指示灯"
   Rectangle "矩形_234" at 75,385 size 44x21
      Appearance <- "输出_5号梯2层按钮指示灯"
   Button "FB_Empty_Rectangular_1" at 82,410 size 29x18; TextOff 'Text'; PictureOff "FB_Empty_Rectangular_Released_256c"; PictureOn "FB_Empty_Rectangular_Pressed_256c"
      on Release: ResetBit("输入_5号梯轿内选层按钮1")
      on Press: SetBit("输入_5号梯轿内选层按钮1")
   Button "FB_Empty_Rectangular_2" at 83,387 size 29x18; TextOff 'Text'; PictureOff "FB_Empty_Rectangular_Released_256c"; PictureOn "FB_Empty_Rectangular_Pressed_256c"
      on Release: ResetBit("输入_5号梯轿内选层按钮2")
      on Press: SetBit("输入_5号梯轿内选层按钮2")
   Rectangle "矩形_235" at 75,363 size 44x21
      Appearance <- "输出_5号梯3层按钮指示灯"
   Button "FB_Empty_Rectangular_3" at 83,365 size 29x18; TextOff 'Text'; PictureOff "FB_Empty_Rectangular_Released_256c"; PictureOn "FB_Empty_Rectangular_Pressed_256c"
      on Release: ResetBit("输入_5号梯轿内选层按钮3")
      on Press: SetBit("输入_5号梯轿内选层按钮3")
   Rectangle "矩形_236" at 75,341 size 44x21
      Appearance <- "输出_5号梯4层按钮指示灯"
   Button "FB_Empty_Rectangular_4" at 83,343 size 29x18; TextOff 'Text'; PictureOff "FB_Empty_Rectangular_Released_256c"; PictureOn "FB_Empty_Rectangular_Pressed_256c"
      on Release: ResetBit("输入_5号梯轿内选层按钮4")
      on Press: SetBit("输入_5号梯轿内选层按钮4")
   Button "FB_Empty_Rectangular_5" at 83,321 size 29x18; TextOff 'Text'; PictureOff "FB_Empty_Rectangular_Released_256c"; PictureOn "FB_Empty_Rectangular_Pressed_256c"
      on Release: ResetBit("输入_5号梯轿内选层按钮5")
      on Press: SetBit("输入_5号梯轿内选层按钮5")
   Button "FB_Empty_Rectangular_6" at 83,299 size 29x18; TextOff 'Text'; PictureOff "FB_Empty_Rectangular_Released_256c"; PictureOn "FB_Empty_Rectangular_Pressed_256c"
      on Release: ResetBit("输入_5号梯轿内选层按钮6")
      on Press: SetBit("输入_5号梯轿内选层按钮6")
   Button "FB_Empty_Rectangular_7" at 83,277 size 29x18; TextOff 'Text'; PictureOff "FB_Empty_Rectangular_Released_256c"; PictureOn "FB_Empty_Rectangular_Pressed_256c"
      on Release: ResetBit("输入_5号梯轿内选层按钮7")
      on Press: SetBit("输入_5号梯轿内选层按钮7")
   Button "FB_Empty_Rectangular_8" at 83,255 size 29x18; TextOff 'Text'; PictureOff "FB_Empty_Rectangular_Released_256c"; PictureOn "FB_Empty_Rectangular_Pressed_256c"
      on Release: ResetBit("输入_5号梯轿内选层按钮8")
      on Press: SetBit("输入_5号梯轿内选层按钮8")
   Button "FB_Empty_Rectangular_9" at 83,233 size 29x18; TextOff 'Text'; PictureOff "FB_Empty_Rectangular_Released_256c"; PictureOn "FB_Empty_Rectangular_Pressed_256c"
      on Release: ResetBit("输入_5号梯轿内选层按钮9")
      on Press: SetBit("输入_5号梯轿内选层按钮9")
   Button "FB_Empty_Rectangular_10" at 83,211 size 29x18; TextOff 'Text'; PictureOff "FB_Empty_Rectangular_Released_256c"; PictureOn "FB_Empty_Rectangular_Pressed_256c"
      on Release: ResetBit("输入_5号梯轿内选层按钮10")
      on Press: SetBit("输入_5号梯轿内选层按钮10")
   TextField "文本域_14" at 90,409 size 14x19; Text '1'
   TextField "文本域_15" at 90,386 size 14x19; Text '2'
   TextField "文本域_16" at 90,363 size 14x19; Text '3'
   TextField "文本域_17" at 90,342 size 14x19; Text '4'
   TextField "文本域_18" at 90,320 size 14x19; Text '5'
   TextField "文本域_19" at 90,298 size 14x19; Text '6'
   TextField "文本域_20" at 90,276 size 14x19; Text '7'
   TextField "文本域_21" at 90,254 size 14x19; Text '8'
   TextField "文本域_22" at 90,232 size 14x19; Text '9'
   TextField "文本域_40" at 86,210 size 23x19; Text '10'
   Circle "圆_56" at 475,117 size 24x24
      Appearance <- "输出_5号梯满载指示"
   Circle "圆_57" at 585,117 size 24x24
      Appearance <- "输出_5号梯故障指示"
   Circle "圆_58" at 473,163 size 24x24
      Appearance <- "输出_5号梯照明指示"
   Circle "圆_59" at 368,122 size 24x24
      Appearance <- "输出_5号梯满载指示"
   Circle "圆_60" at 584,165 size 24x24
      Appearance <- "输出_5号梯风扇指示"
   TextField "文本域_47" at 402,119 size 45x23; Text '超重'
   TextField "文本域_48" at 509,120 size 45x23; Text '满载'
   TextField "文本域_49" at 621,119 size 45x23; Text '故障'
   TextField "文本域_50" at 511,166 size 45x23; Text '照明'
   TextField "文本域_51" at 621,166 size 45x23; Text '风扇'
   Circle "圆_73" at 226,119 size 24x24
      Appearance <- "输入_自动运行信号"
   TextField "文本域_68" at 257,120 size 73x20; Text '自动运行'
   TextField "文本域_69" at 256,167 size 107x20; Text '电梯准备就绪'
   Circle "圆_83" at 473,348 size 16x16
      Appearance <- "输出_5号梯开门继电器"
   Circle "圆_86" at 473,363 size 16x16
      Appearance <- "输出_5号梯关门继电器"
   Circle "圆_89" at 630,264 size 16x16
      Appearance <- "输入_5号梯开门到位"
   Circle "圆_92" at 630,280 size 16x16
      Appearance <- "输入_5号梯关门到位"
   Circle "圆_129" at 630,212 size 16x16
      Appearance <- "输出_5号梯电机启动信号"
   Circle "圆_132" at 630,227 size 16x16
      Appearance <- "输出_5号梯上行接触器"
   Circle "圆_135" at 630,242 size 16x16
      Appearance <- "输出_5号梯下行接触器"
   Circle "圆_19" at 226,163 size 24x24
      Appearance <- "输出_准备就绪信号"
   Circle "圆_95" at 630,335 size 16x16
      Appearance <- "输出_5号梯1级减速制动"
   Circle "圆_98" at 630,350 size 16x16
      Appearance <- "输出_5号梯2级减速制动"
   Circle "圆_101" at 630,365 size 16x16
      Appearance <- "输出_5号梯3级减速制动"
   Circle "圆_104" at 630,304 size 16x16
      Appearance <- "输出_5号梯低速接触器"
   Circle "圆_107" at 630,319 size 16x16
      Appearance <- "输出_5号梯高速接触器"
   Circle "圆_120" at 330,365 size 16x16
      Appearance <- "输入_5号梯轿厢门锁信号"
   Circle "圆_123" at 330,214 size 16x16
      Appearance <- "输入_5号梯10楼层门锁信号"
   Circle "圆_126" at 330,229 size 16x16
      Appearance <- "输入_5号梯9楼层门锁信号"
   Circle "圆_138" at 330,244 size 16x16
      Appearance <- "输入_5号梯8楼层门锁信号"
   Circle "圆_141" at 330,259 size 16x16
      Appearance <- "输入_5号梯7楼层门锁信号"
   Circle "圆_144" at 330,274 size 16x16
      Appearance <- "输入_5号梯6楼层门锁信号"
   Circle "圆_147" at 330,289 size 16x16
      Appearance <- "输入_1号梯5楼层门锁信号"
   Circle "圆_150" at 330,304 size 16x16
      Appearance <- "输入_5号梯4楼层门锁信号"
   Circle "圆_153" at 330,319 size 16x16
      Appearance <- "输入_5号梯3楼层门锁信号"
   Circle "圆_156" at 330,334 size 16x16
      Appearance <- "输入_5号梯2楼层门锁信号"
   Circle "圆_159" at 330,349 size 16x16
      Appearance <- "输入_5号梯1楼层门锁信号"
   Circle "圆_162" at 474,213 size 16x16
      Appearance <- "输入_5号梯上端站第2限位"
   Circle "圆_165" at 474,228 size 16x16
      Appearance <- "输入_5号梯上端站第1限位"
   Circle "圆_168" at 474,243 size 16x16
      Appearance <- "输入_5号梯上平层信号"
   Circle "圆_171" at 474,258 size 16x16
      Appearance <- "输入_5号梯下平层信号"
   Circle "圆_174" at 474,273 size 16x16
      Appearance <- "输入_5号梯下端站第2限位"
   Circle "圆_177" at 474,288 size 16x16
      Appearance <- "输入_5号梯下端站第1限位"
   Circle "圆_183" at 474,315 size 16x16
      Appearance <- "输入_5号梯检修信号"
   Circle "圆_186" at 474,330 size 16x16
      Appearance <- "输入_5号梯光幕信号"
   Rectangle "矩形_193" at 167,134 size 4x18
      Appearance <- "输出_5号梯LEDi"
   Rectangle "矩形_194" at 167,156 size 4x18
      Appearance <- "输出_5号梯LEDj"
   Rectangle "矩形_195" at 180,132 size 18x4
      Appearance <- "输出_5号梯LEDa"
   Rectangle "矩形_196" at 177,136 size 4x18
      Appearance <- "输出_5号梯LEDf"
   Rectangle "矩形_197" at 180,153 size 18x4
      Appearance <- "输出_5号梯LEDg"
   Rectangle "矩形_198" at 177,157 size 4x18
      Appearance <- "输出_5号梯LEDe"
   Rectangle "矩形_199" at 180,175 size 18x4
      Appearance <- "输出_5号梯LEDd"
   Rectangle "矩形_200" at 197,135 size 4x18
      Appearance <- "输出_5号梯LEDb"
   Rectangle "矩形_201" at 197,157 size 4x18
      Appearance <- "输出_5号梯LEDc"
   Rectangle "矩形_72" at 93,122 size 6x34
      Appearance <- "输出_5号梯上行指示"
   Polygon "多边形_5" at 81,118 size 15x17
      Appearance <- "输出_5号梯上行指示"
   Polygon "多边形_6" at 96,118 size 14x17
      Appearance <- "输出_5号梯上行指示"
   Rectangle "矩形_73" at 93,157 size 6x34
      Appearance <- "输出_5号梯下行指示"
   Polygon "多边形_1" at 79,179 size 17x15
      Appearance <- "输出_5号梯下行指示"
   Polygon "多边形_2" at 96,179 size 17x15
      Appearance <- "输出_5号梯下行指示"
   TextField "文本域_77" at 225,230 size 81x15; Text '9层门锁信号'
   TextField "文本域_78" at 225,244 size 81x15; Text '8层门锁信号'
   TextField "文本域_79" at 225,259 size 81x15; Text '7层门锁信号'
   TextField "文本域_80" at 225,274 size 81x15; Text '6层门锁信号'
   TextField "文本域_81" at 225,289 size 81x15; Text '5层门锁信号'
   TextField "文本域_83" at 225,304 size 81x15; Text '4层门锁信号'
   TextField "文本域_84" at 225,319 size 81x15; Text '3层门锁信号'
   TextField "文本域_85" at 225,336 size 81x15; Text '2层门锁信号'
   TextField "文本域_86" at 224,352 size 82x15; Text '1层门锁信号'
   TextField "文本域_87" at 220,367 size 86x15; Text '轿厢门锁信号'
   TextField "文本域_23" at 395,312 size 72x15; Text '检修开关'
   TextField "文本域_24" at 397,328 size 70x15; Text '光幕信号'
   TextField "文本域_82" at 364,215 size 103x15; Text '上端站第二限位'
   TextField "文本域_88" at 363,231 size 104x15; Text '上端站第一限位'
   TextField "文本域_89" at 385,246 size 82x15; Text '上平层信号'
   TextField "文本域_90" at 385,261 size 82x15; Text '下平层信号'
   TextField "文本域_91" at 363,275 size 104x15; Text '下端站第二限位'
   TextField "文本域_92" at 363,291 size 104x15; Text '下端站第一限位'
   TextField "文本域_13" at 375,348 size 93x15; Text '开门到位信号'
   TextField "文本域_25" at 375,364 size 93x15; Text '关门到位信号'
   TextField "文本域_97" at 529,267 size 92x15; Text '开门继电器'
   TextField "文本域_98" at 529,283 size 92x15; Text '关门继电器'
   TextField "文本域_104" at 529,249 size 92x15; Text '下行接触器'
   TextField "文本域_105" at 518,217 size 103x15; Text '电机启动信号'
   TextField "文本域_106" at 529,233 size 92x15; Text '上行接触器'
   TextField "文本域_99" at 508,351 size 114x15; Text '二级制动接触器'
   TextField "文本域_100" at 508,367 size 114x15; Text '三级制动接触器'
   TextField "文本域_101" at 508,334 size 114x15; Text '一级制动接触器'
   TextField "文本域_102" at 508,302 size 114x15; Text '低速运行接触器'
   TextField "文本域_103" at 508,318 size 114x15; Text '高速运行接触器'
   TextField "文本域_76" at 219,214 size 91x15; Text '10层门锁信号'
   Clock "时钟_1" at 664,57 size 101x57
   DateTimeField "日期/时间域_1" at 491,71 size 184x28
   TextField "文本域_26" at 260,403 size 142x19; Text '1号电梯开关门状态'
   Button "FB_Left_Square" at 284,442 size 20x20; TextOff 'Text'; PictureOff "FB_Left_Square_Released_256c"; PictureOn "FB_Left_Square_Pressed_256c"
      on Click: SetBit("输入_1号梯轿内开门按钮")
      Appearance <- "输入_5号梯轿内开门按钮"
   Button "FB_Right_Square" at 304,442 size 20x20; TextOff 'Text'; PictureOff "FB_Right_Square_Released_256c_5"; PictureOn "FB_Right_Square_Pressed_256c"
      on Click: SetBit("输入_1号梯轿内开门按钮")
      Appearance <- "输入_1号梯轿内开门按钮"
   Button "FB_Left_Square_1" at 350,442 size 20x20; TextOff 'Text'; PictureOff "FB_Left_Square_Released_256c"; PictureOn "FB_Left_Square_Pressed_256c"
      on Click: SetBit("输入_1号梯轿内关门按钮")
      Appearance <- "输入_5号梯轿内关门按钮"
   Button "FB_Right_Square_1" at 330,442 size 20x20; TextOff 'Text'; PictureOff "FB_Right_Square_Released_256c_5"; PictureOn "FB_Right_Square_Pressed_256c"
      on Click: SetBit("输入_1号梯轿内关门按钮")
      Appearance <- "输入_1号梯轿内关门按钮"

screen "6#电梯状态画面" 800x600
   TextField "文本域_1" at 385,17 size 280x27; Text '-- 6#电梯状态总览'
   TextField "文本域_3" at 69,12 size 308x31; Text '电 梯 监 控 系 统'
   Button "按钮_7" at 557,519 size 117x65; TextOff '电梯状态总览'
      on Click: ActivateScreen("电梯状态总览画面", 0)
   Button "按钮_8" at 680,518 size 106x65; TextOff '退出系统'
      on Click: StopRuntime(0)
   Group "Group" at 290,421 size 40x20; PictureOn "FB_Left_Square_Pressed_256c"; PictureOff "FB_Left_Square_Released_256c"
   Group "Group_1" at 337,420 size 40x20; PictureOn "FB_Left_Square_Pressed_256c"; PictureOff "FB_Left_Square_Released_256c"
   Rectangle "矩形_237" at 74,311 size 44x21
      Appearance <- "输出_1号梯5层按钮指示灯"
   Rectangle "矩形_238" at 74,289 size 44x21
      Appearance <- "输出_1号梯6层按钮指示灯"
   Rectangle "矩形_239" at 74,267 size 44x21
      Appearance <- "输出_1号梯7层按钮指示灯"
   Rectangle "矩形_240" at 74,245 size 44x21
      Appearance <- "输出_1号梯8层按钮指示灯"
   Rectangle "矩形_241" at 74,223 size 44x21
      Appearance <- "输出_1号梯9层按钮指示灯"
   Rectangle "矩形_242" at 74,201 size 44x21
      Appearance <- "输出_1号梯10层按钮指示灯"
   Circle "圆_1" at 162,204 size 14x14
      Appearance <- "输出_10层下行呼梯按钮指示灯"
   Circle "圆_2" at 150,226 size 14x14
      Appearance <- "输出_9层上行呼梯按钮指示灯"
   Circle "圆_3" at 175,226 size 14x14
      Appearance <- "输出_9层下行呼梯按钮指示灯"
   Circle "圆_4" at 150,249 size 14x14
      Appearance <- "输出_8层上行呼梯按钮指示灯"
   Circle "圆_5" at 175,249 size 14x14
      Appearance <- "输出_8层下行呼梯按钮指示灯"
   Circle "圆_6" at 150,269 size 14x14
      Appearance <- "输出_7层上行呼梯按钮指示灯"
   Circle "圆_7" at 175,269 size 14x14
      Appearance <- "输出_7层下行呼梯按钮指示灯"
   Circle "圆_8" at 150,291 size 14x14
      Appearance <- "输出_6层上行呼梯按钮指示灯"
   Circle "圆_9" at 175,291 size 14x14
      Appearance <- "输出_6层下行呼梯按钮指示灯"
   Circle "圆_10" at 150,314 size 14x14
      Appearance <- "输出_5层上行呼梯按钮指示灯"
   Circle "圆_11" at 175,314 size 14x14
      Appearance <- "输出_5层下行呼梯按钮指示灯"
   Circle "圆_12" at 150,336 size 14x14
      Appearance <- "输出_4层上行呼梯按钮指示灯"
   Circle "圆_13" at 175,336 size 14x14
      Appearance <- "输出_4层下行呼梯按钮指示灯"
   Circle "圆_14" at 150,360 size 14x14
      Appearance <- "输出_3层上行呼梯按钮指示灯"
   Circle "圆_15" at 175,360 size 14x14
      Appearance <- "输出_3层下行呼梯按钮指示灯"
   Circle "圆_16" at 150,381 size 14x14
      Appearance <- "输出_2层上行呼梯按钮指示灯"
   Circle "圆_17" at 175,381 size 14x14
      Appearance <- "输出_2层下行呼梯按钮指示灯"
   Circle "圆_18" at 163,404 size 14x14
      Appearance <- "输出_1层上行呼梯按钮指示灯"
   TextField "文本域_41" at 76,432 size 45x23; Text '内呼'
   TextField "文本域_42" at 155,432 size 45x23; Text '外呼'
   Rectangle "矩形_233" at 74,399 size 44x21
      Appearance <- "输出_1号梯1层按钮指示灯"
   Rectangle "矩形_234" at 74,377 size 44x21
      Appearance <- "输出_1号梯2层按钮指示灯"
   Button "FB_Empty_Rectangular_1" at 81,402 size 29x18; TextOff 'Text'; PictureOff "FB_Empty_Rectangular_Released_256c"; PictureOn "FB_Empty_Rectangular_Pressed_256c"
      on Release: ResetBit("输入_1号梯轿内选层按钮1")
      on Press: SetBit("输入_1号梯轿内选层按钮1")
      Appearance <- "输出_1号梯1层按钮指示灯"
   Button "FB_Empty_Rectangular_2" at 82,379 size 29x18; TextOff 'Text'; PictureOff "FB_Empty_Rectangular_Released_256c"; PictureOn "FB_Empty_Rectangular_Pressed_256c"
      on Release: ResetBit("输入_1号梯轿内选层按钮2")
      on Press: SetBit("输入_1号梯轿内选层按钮2")
   Rectangle "矩形_235" at 74,355 size 44x21
      Appearance <- "输出_1号梯3层按钮指示灯"
   Button "FB_Empty_Rectangular_3" at 82,357 size 29x18; TextOff 'Text'; PictureOff "FB_Empty_Rectangular_Released_256c"; PictureOn "FB_Empty_Rectangular_Pressed_256c"
      on Release: ResetBit("输入_1号梯轿内选层按钮3")
      on Press: SetBit("输入_1号梯轿内选层按钮3")
   Rectangle "矩形_236" at 74,333 size 44x21
      Appearance <- "输出_1号梯4层按钮指示灯"
   Button "FB_Empty_Rectangular_4" at 82,335 size 29x18; TextOff 'Text'; PictureOff "FB_Empty_Rectangular_Released_256c"; PictureOn "FB_Empty_Rectangular_Pressed_256c"
      on Release: ResetBit("输入_1号梯轿内选层按钮4")
      on Press: SetBit("输入_1号梯轿内选层按钮4")
   Button "FB_Empty_Rectangular_5" at 82,313 size 29x18; TextOff 'Text'; PictureOff "FB_Empty_Rectangular_Released_256c"; PictureOn "FB_Empty_Rectangular_Pressed_256c"
      on Release: ResetBit("输入_1号梯轿内选层按钮5")
      on Press: SetBit("输入_1号梯轿内选层按钮5")
   Button "FB_Empty_Rectangular_6" at 82,291 size 29x18; TextOff 'Text'; PictureOff "FB_Empty_Rectangular_Released_256c"; PictureOn "FB_Empty_Rectangular_Pressed_256c"
      on Release: ResetBit("输入_1号梯轿内选层按钮6")
      on Press: SetBit("输入_1号梯轿内选层按钮6")
   Button "FB_Empty_Rectangular_7" at 82,269 size 29x18; TextOff 'Text'; PictureOff "FB_Empty_Rectangular_Released_256c"; PictureOn "FB_Empty_Rectangular_Pressed_256c"
      on Release: ResetBit("输入_1号梯轿内选层按钮7")
      on Press: SetBit("输入_1号梯轿内选层按钮7")
   Button "FB_Empty_Rectangular_8" at 82,247 size 29x18; TextOff 'Text'; PictureOff "FB_Empty_Rectangular_Released_256c"; PictureOn "FB_Empty_Rectangular_Pressed_256c"
      on Release: ResetBit("输入_1号梯轿内选层按钮8")
      on Press: SetBit("输入_1号梯轿内选层按钮8")
   Button "FB_Empty_Rectangular_9" at 82,225 size 29x18; TextOff 'Text'; PictureOff "FB_Empty_Rectangular_Released_256c"; PictureOn "FB_Empty_Rectangular_Pressed_256c"
      on Release: ResetBit("输入_1号梯轿内选层按钮9")
      on Press: SetBit("输入_1号梯轿内选层按钮9")
   Button "FB_Empty_Rectangular_10" at 82,203 size 29x18; TextOff 'Text'; PictureOff "FB_Empty_Rectangular_Released_256c"; PictureOn "FB_Empty_Rectangular_Pressed_256c"
      on Release: ResetBit("输入_1号梯轿内选层按钮10")
      on Press: SetBit("输入_1号梯轿内选层按钮10")
   TextField "文本域_14" at 89,401 size 14x19; Text '1'
   TextField "文本域_15" at 89,378 size 14x19; Text '2'
   TextField "文本域_16" at 89,355 size 14x19; Text '3'
   TextField "文本域_17" at 89,334 size 14x19; Text '4'
   TextField "文本域_18" at 89,312 size 14x19; Text '5'
   TextField "文本域_19" at 89,290 size 14x19; Text '6'
   TextField "文本域_20" at 89,268 size 14x19; Text '7'
   TextField "文本域_21" at 89,246 size 14x19; Text '8'
   TextField "文本域_22" at 89,224 size 14x19; Text '9'
   TextField "文本域_40" at 85,202 size 23x19; Text '10'
   Circle "圆_56" at 471,111 size 24x24
      Appearance <- "输出_6号梯满载指示"
   Circle "圆_57" at 581,111 size 24x24
      Appearance <- "输出_6号梯故障指示"
   Circle "圆_58" at 470,160 size 24x24
      Appearance <- "输出_6号梯照明指示"
   Circle "圆_59" at 370,113 size 24x24
      Appearance <- "输出_6号梯满载指示"
   Circle "圆_60" at 581,162 size 24x24
      Appearance <- "输出_6号梯风扇指示"
   TextField "文本域_47" at 399,112 size 45x23; Text '超重'
   TextField "文本域_48" at 505,114 size 45x23; Text '满载'
   TextField "文本域_49" at 617,113 size 45x23; Text '故障'
   TextField "文本域_50" at 508,163 size 45x23; Text '照明'
   TextField "文本域_51" at 618,163 size 45x23; Text '风扇'
   Circle "圆_73" at 223,112 size 24x24
      Appearance <- "输入_自动运行信号"
   TextField "文本域_68" at 254,113 size 73x20; Text '自动运行'
   TextField "文本域_69" at 253,160 size 107x20; Text '电梯准备就绪'
   Circle "圆_83" at 471,339 size 16x16
      Appearance <- "输出_6号梯开门继电器"
   Circle "圆_86" at 471,354 size 16x16
      Appearance <- "输出_6号梯关门继电器"
   Circle "圆_89" at 627,259 size 16x16
      Appearance <- "输入_6号梯开门到位"
   Circle "圆_92" at 627,275 size 16x16
      Appearance <- "输入_6号梯关门到位"
   Circle "圆_129" at 627,208 size 16x16
      Appearance <- "输出_6号梯电机启动信号"
   Circle "圆_132" at 627,223 size 16x16
      Appearance <- "输出_6号梯上行指示"
   Circle "圆_135" at 627,238 size 16x16
      Appearance <- "输出_6号梯下行指示"
   Circle "圆_19" at 223,156 size 24x24
      Appearance <- "输出_准备就绪信号"
   Circle "圆_95" at 627,330 size 16x16
      Appearance <- "输出_6号梯1级减速制动"
   Circle "圆_98" at 627,345 size 16x16
      Appearance <- "输出_6号梯2级减速制动"
   Circle "圆_101" at 627,360 size 16x16
      Appearance <- "输出_6号梯3级减速制动"
   Circle "圆_104" at 627,299 size 16x16
      Appearance <- "输出_6号梯低速接触器"
   Circle "圆_107" at 627,314 size 16x16
      Appearance <- "输出_6号梯高速接触器"
   Circle "圆_120" at 320,361 size 16x16
      Appearance <- "输入_6号梯轿厢门锁信号"
   Circle "圆_123" at 320,210 size 16x16
      Appearance <- "输入_6号梯10楼层门锁信号"
   Circle "圆_126" at 320,225 size 16x16
      Appearance <- "输入_6号梯9楼层门锁信号"
   Circle "圆_138" at 320,240 size 16x16
      Appearance <- "输入_6号梯8楼层门锁信号"
   Circle "圆_141" at 320,255 size 16x16
      Appearance <- "输入_6号梯7楼层门锁信号"
   Circle "圆_144" at 320,270 size 16x16
      Appearance <- "输入_6号梯6楼层门锁信号"
   Circle "圆_147" at 320,285 size 16x16
      Appearance <- "输入_6号梯5楼层门锁信号"
   Circle "圆_150" at 320,300 size 16x16
      Appearance <- "输入_6号梯4楼层门锁信号"
   Circle "圆_153" at 320,315 size 16x16
      Appearance <- "输入_6号梯3楼层门锁信号"
   Circle "圆_156" at 320,330 size 16x16
      Appearance <- "输入_6号梯2楼层门锁信号"
   Circle "圆_159" at 320,345 size 16x16
      Appearance <- "输入_6号梯1楼层门锁信号"
   Circle "圆_162" at 471,210 size 16x16
      Appearance <- "输入_6号梯上端站第2限位"
   Circle "圆_165" at 471,225 size 16x16
      Appearance <- "输入_6号梯上端站第1限位"
   Circle "圆_168" at 471,240 size 16x16
      Appearance <- "输入_6号梯上平层信号"
   Circle "圆_171" at 471,255 size 16x16
      Appearance <- "输入_6号梯下平层信号"
   Circle "圆_174" at 471,270 size 16x16
      Appearance <- "输入_6号梯下端站第2限位"
   Circle "圆_177" at 471,285 size 16x16
      Appearance <- "输入_6号梯下端站第1限位"
   Circle "圆_183" at 471,306 size 16x16
      Appearance <- "输入_6号梯检修信号"
   Circle "圆_186" at 471,321 size 16x16
      Appearance <- "输入_6号梯光幕信号"
   Rectangle "矩形_193" at 166,126 size 4x18
      Appearance <- "输出_6号梯LEDi"
   Rectangle "矩形_194" at 166,148 size 4x18
      Appearance <- "输出_6号梯LEDj"
   Rectangle "矩形_195" at 179,124 size 18x4
      Appearance <- "输出_6号梯LEDa"
   Rectangle "矩形_196" at 176,128 size 4x18
      Appearance <- "输出_6号梯LEDf"
   Rectangle "矩形_197" at 179,145 size 18x4
      Appearance <- "输出_6号梯LEDg"
   Rectangle "矩形_198" at 176,149 size 4x18
      Appearance <- "输出_6号梯LEDe"
   Rectangle "矩形_199" at 179,167 size 18x4
      Appearance <- "输出_6号梯LEDd"
   Rectangle "矩形_200" at 196,127 size 4x18
      Appearance <- "输出_6号梯LEDb"
   Rectangle "矩形_201" at 196,149 size 4x18
      Appearance <- "输出_6号梯LEDc"
   Rectangle "矩形_72" at 92,114 size 6x34
      Appearance <- "输出_6号梯上行指示"
   Polygon "多边形_5" at 80,110 size 15x17
      Appearance <- "输出_6号梯上行指示"
   Polygon "多边形_6" at 95,110 size 14x17
      Appearance <- "输出_6号梯上行指示"
   Rectangle "矩形_73" at 92,149 size 6x34
      Appearance <- "输出_6号梯下行指示"
   Polygon "多边形_1" at 78,171 size 17x15
      Appearance <- "输出_6号梯下行指示"
   Polygon "多边形_2" at 95,171 size 17x15
      Appearance <- "输出_6号梯下行指示"
   TextField "文本域_77" at 224,227 size 81x15; Text '9层门锁信号'
   TextField "文本域_78" at 224,241 size 81x15; Text '8层门锁信号'
   TextField "文本域_79" at 224,256 size 81x15; Text '7层门锁信号'
   TextField "文本域_80" at 224,271 size 81x15; Text '6层门锁信号'
   TextField "文本域_81" at 224,286 size 81x15; Text '5层门锁信号'
   TextField "文本域_83" at 224,301 size 81x15; Text '4层门锁信号'
   TextField "文本域_84" at 224,316 size 81x15; Text '3层门锁信号'
   TextField "文本域_85" at 224,331 size 81x15; Text '2层门锁信号'
   TextField "文本域_86" at 223,347 size 82x15; Text '1层门锁信号'
   TextField "文本域_87" at 224,361 size 81x15; Text '轿厢门锁信号'
   TextField "文本域_23" at 388,305 size 72x15; Text '检修开关'
   TextField "文本域_24" at 390,321 size 70x15; Text '光幕信号'
   TextField "文本域_82" at 357,212 size 103x15; Text '上端站第二限位'
   TextField "文本域_88" at 356,228 size 104x15; Text '上端站第一限位'
   TextField "文本域_89" at 378,243 size 82x15; Text '上平层信号'
   TextField "文本域_90" at 378,258 size 82x15; Text '下平层信号'
   TextField "文本域_91" at 356,272 size 104x15; Text '下端站第二限位'
   TextField "文本域_92" at 356,288 size 104x15; Text '下端站第一限位'
   TextField "文本域_13" at 368,342 size 93x15; Text '开门到位信号'
   TextField "文本域_25" at 368,358 size 93x15; Text '关门到位信号'
   TextField "文本域_97" at 528,262 size 92x15; Text '开门继电器'
   TextField "文本域_98" at 528,278 size 92x15; Text '关门继电器'
   TextField "文本域_104" at 528,243 size 92x15; Text '下行接触器'
   TextField "文本域_105" at 517,211 size 103x15; Text '电机启动信号'
   TextField "文本域_106" at 528,227 size 92x15; Text '上行接触器'
   TextField "文本域_99" at 507,347 size 114x15; Text '二级制动接触器'
   TextField "文本域_100" at 507,363 size 114x15; Text '三级制动接触器'
   TextField "文本域_101" at 507,330 size 114x15; Text '一级制动接触器'
   TextField "文本域_102" at 507,298 size 114x15; Text '低速运行接触器'
   TextField "文本域_103" at 507,314 size 114x15; Text '高速运行接触器'
   TextField "文本域_76" at 218,212 size 91x15; Text '10层门锁信号'
   Clock "时钟_1" at 664,57 size 101x57
   DateTimeField "日期/时间域_1" at 491,71 size 184x28
   TextField "文本域_26" at 257,385 size 142x19; Text '1号电梯开关门状态'
   Button "FB_Left_Square" at 290,421 size 20x20; TextOff 'Text'; PictureOff "FB_Left_Square_Released_256c"; PictureOn "FB_Left_Square_Pressed_256c"
      on Click: SetBit("输入_6号梯轿内开门按钮")
      Appearance <- "输入_1号梯轿内开门按钮"
   Button "FB_Right_Square" at 310,421 size 20x20; TextOff 'Text'; PictureOff "FB_Right_Square_Released_256c_6"; PictureOn "FB_Right_Square_Pressed_256c"
      on Click: SetBit("输入_1号梯轿内开门按钮")
      Appearance <- "输入_1号梯轿内开门按钮"
   Button "FB_Left_Square_1" at 357,420 size 20x20; TextOff 'Text'; PictureOff "FB_Left_Square_Released_256c"; PictureOn "FB_Left_Square_Pressed_256c"
      on Click: SetBit("输入_1号梯轿内关门按钮")
      Appearance <- "输入_1号梯轿内关门按钮"
   Button "FB_Right_Square_1" at 337,420 size 20x20; TextOff 'Text'; PictureOff "FB_Right_Square_Released_256c_6"; PictureOn "FB_Right_Square_Pressed_256c"
      on Click: SetBit("输入_1号梯轿内关门按钮")
      Appearance <- "输入_1号梯轿内关门按钮"

screen "主画面" 800x600
   TextField "文本域_1" at 294,117 size 85x35; Text '，欢迎您！'
   TextField "文本域_2" at 192,169 size 103x32; Text '您的身份是：'
   IOField "I/O 域_1" at 189,110 size 99x32; FormatPattern ????????????????????????????????????????????????????????????????????????????????
      ProcessValue <- "用户名"
   Button "按钮_2" at 490,152 size 166x42; TextOff '电梯运行监控'
      on Click: ActivateScreen("电梯运行监控画面1", 0)
   Button "按钮_3" at 490,200 size 166x42; TextOff '外呼状态监控'
      on Click: ActivateScreen("外呼状态监控画面", 0)
   Button "按钮_4" at 491,296 size 166x42; TextOff '设置'; Authorization "监视"
      on Click: ActivateScreen("设置画面", 0)
      Visibility <- "zuhao"
   Button "按钮_5" at 490,344 size 166x42; TextOff '注销'
      on Click: function_f23ef4c9(); ActivateScreen("登录画面", 0)
   Button "按钮_6" at 491,248 size 166x42; TextOff '电梯状态记录'
      on Click: ActivateScreen("运行数据记录", 0)
      Visibility <- "zuhao"
   SymbolicIOField "符号 I/O 域_1" at 294,162 size 72x32; TextOn '管理员'; TextOff '0'; TextList "身份"
   Button "按钮_7" at 564,517 size 110x66; TextOff '登录画面'
      on Click: ActivateScreen("登录画面", 0)
   TextField "文本域_3" at 241,11 size 323x31; Text '电 梯 监 控 系 统'
   Button "按钮_8" at 682,517 size 106x66; TextOff '退出系统'
      on Click: StopRuntime(0)
   Button "按钮_9" at 490,104 size 166x42; TextOff '电梯状态总览'
      on Click: ActivateScreen("电梯状态总览画面", 0)
   Clock "时钟_1" at 664,57 size 101x57
   DateTimeField "日期/时间域_1" at 491,71 size 184x28
   TextField "文本域_4" at 117,230 size 126x17; Text '电梯名称：CIMC-EET'
   TextField "文本域_5" at 117,247 size 133x17; Text '电梯编号：CIMC-2023'
   TextField "文本域_6" at 117,264 size 124x17; Text '维保单位：CIMC大学'
   TextField "文本域_7" at 115,296 size 57x17; Text '当前状态'
   TextField "文本域_8" at 117,318 size 83x17; Text '控制器状态：'
   TextField "文本域_9" at 114,346 size 70x17; Text '工作状态：'
   TextField "文本域_10" at 115,385 size 96x17; Text '当前运行时间：'
   TextField "文本域_11" at 200,315 size 37x19; Text '在线'
      Visibility <- "输入_自动运行信号"
   TextField "文本域_12" at 202,315 size 37x19; Text '离线'
      Visibility <- "输入_自动运行信号"
   TextField "文本域_13" at 186,345 size 53x19; Text '初始化'
      Visibility <- "输入_自动运行信号"
   TextField "文本域_15" at 189,344 size 69x19; Text '正在接客'
      Visibility <- "输出_准备就绪信号"
   IOField "I/O 域_2" at 211,378 size 35x32; FormatPattern 99
      ProcessValue <- "程序运行小时"
   TextField "文本域_14" at 246,379 size 20x31; Text ':'
   IOField "I/O 域_3" at 269,378 size 35x32; FormatPattern 99
      ProcessValue <- "程序运行分钟"
   TextField "文本域_16" at 304,379 size 20x31; Text ':'
   IOField "I/O 域_4" at 324,378 size 35x32; FormatPattern 99
      ProcessValue <- "程序运行秒"

screen "初始化楼层设定" 800x600
   Button "按钮_7" at 560,516 size 110x66; TextOff '主画面'
      on Click: ActivateScreen("主画面", 0)
   TextField "文本域_1" at 385,17 size 280x27; Text '-- 初始化楼层设定'
   TextField "文本域_3" at 91,12 size 286x31; Text '电 梯 监 控 系 统'
   Button "按钮_1" at 676,516 size 106x66; TextOff '退出系统'
      on Click: StopRuntime(0)
   IOField "I/O 域_1" at 220,111 size 95x34; FormatPattern s99999
      ProcessValue <- "初始化设置用_1号梯初始化楼层赋值"
   IOField "I/O 域_3" at 220,167 size 95x34; FormatPattern s99999
      ProcessValue <- "初始化设置用_2号梯初始化楼层赋值"
   IOField "I/O 域_5" at 220,227 size 95x34; FormatPattern s99999
      ProcessValue <- "初始化设置用_3号梯初始化楼层赋值"
   IOField "I/O 域_7" at 220,297 size 95x34; FormatPattern s99999
      ProcessValue <- "初始化设置用_4号梯初始化楼层赋值"
   IOField "I/O 域_9" at 220,352 size 95x34; FormatPattern s99999
      ProcessValue <- "初始化设置用_5号梯初始化楼层赋值"
   IOField "I/O 域_11" at 220,417 size 95x34; FormatPattern s99999
      ProcessValue <- "初始化设置用_6号梯初始化楼层赋值"
   TextField "文本域_2" at 70,106 size 148x40; Text '1#初始化楼层：'
   TextField "文本域_4" at 70,168 size 140x38; Text '2#初始化楼层：'
   TextField "文本域_5" at 70,224 size 139x39; Text '3#初始化楼层：'
   TextField "文本域_6" at 70,298 size 144x36; Text '4#初始化楼层：'
   TextField "文本域_7" at 70,353 size 140x41; Text '5#初始化楼层：'
   TextField "文本域_8" at 70,416 size 144x39; Text '6#初始化楼层：'
   Clock "时钟_1" at 664,57 size 101x57
   DateTimeField "日期/时间域_1" at 491,71 size 184x28
   TextField "文本域_9" at 350,106 size 235x40; Text '1#初始化方向：'
   TextField "文本域_10" at 350,168 size 235x40; Text '2#初始化方向：'
   TextField "文本域_11" at 350,230 size 235x40; Text '3#初始化方向：'
   TextField "文本域_12" at 350,292 size 235x40; Text '4#初始化方向：'
   TextField "文本域_13" at 350,354 size 235x40; Text '5#初始化方向：'
   TextField "文本域_14" at 350,416 size 235x40; Text '6#初始化方向：'
   Switch "开关_1" at 502,97 size 97x44; TextOn '上行'; CaptionText 'Switch'; TextOff '下行'
      ProcessValue <- "初始化设置用_1号梯初始化方向选择"
   Switch "开关_2" at 502,159 size 97x44; TextOn '上行'; CaptionText 'Switch'; TextOff '下行'
      ProcessValue <- "初始化设置用_2号梯初始化方向选择"
   Switch "开关_3" at 502,220 size 97x44; TextOn '上行'; CaptionText 'Switch'; TextOff '下行'
      ProcessValue <- "初始化设置用_3号梯初始化方向选择"
   Switch "开关_4" at 502,283 size 97x44; TextOn '上行'; CaptionText 'Switch'; TextOff '下行'
      ProcessValue <- "初始化设置用_4号梯初始化方向选择"
   Switch "开关_5" at 502,344 size 97x44; TextOn '上行'; CaptionText 'Switch'; TextOff '下行'
      ProcessValue <- "初始化设置用_5号梯初始化方向选择"
   Switch "开关_6" at 502,406 size 97x44; TextOn '上行'; CaptionText 'Switch'; TextOff '下行'
      ProcessValue <- "初始化设置用_6号梯初始化方向选择"

screen "外呼状态监控画面" 800x600
   Button "按钮_7" at 563,519 size 110x66; TextOff '主画面'
      on Click: ActivateScreen("主画面", 0)
   TextField "文本域_1" at 385,17 size 319x27; Text '-- 电梯外呼状态监控'
   TextField "文本域_3" at 114,12 size 263x31; Text '电 梯 监 控 系 统'
   Button "按钮_1" at 682,518 size 106x66; TextOff '退出系统'
      on Click: StopRuntime(0)
   TextField "文本域_2" at 222,83 size 45x19; Text '10F'
   TextField "文本域_4" at 227,124 size 36x19; Text '9F'
   TextField "文本域_5" at 227,176 size 32x19; Text '8F'
   TextField "文本域_6" at 225,225 size 36x19; Text '7F'
   TextField "文本域_7" at 227,273 size 35x19; Text '6F'
   TextField "文本域_8" at 226,372 size 34x19; Text '4F'
   TextField "文本域_9" at 225,323 size 35x19; Text '5F'
   TextField "文本域_10" at 226,421 size 32x19; Text '3F'
   TextField "文本域_11" at 226,470 size 35x19; Text '2F'
   TextField "文本域_12" at 226,510 size 32x19; Text '1F'
   TextField "文本域_13" at 374,116 size 67x19; Text '1#电梯'
   TextField "文本域_14" at 516,115 size 68x19; Text '2#电梯'
   TextField "文本域_15" at 380,253 size 62x19; Text '3#电梯'
   TextField "文本域_16" at 525,253 size 62x19; Text '4#电梯'
   TextField "文本域_17" at 379,392 size 64x19; Text '5#电梯'
   TextField "文本域_18" at 516,392 size 65x19; Text '6#电梯'
   Rectangle "矩形_193" at 414,167 size 4x18
      Appearance <- "输出_1号梯LEDi"
   Rectangle "矩形_194" at 414,189 size 4x18
      Appearance <- "输出_1号梯LEDj"
   Rectangle "矩形_195" at 427,165 size 18x4
      Appearance <- "输出_1号梯LEDa"
   Rectangle "矩形_196" at 424,169 size 4x18
      Appearance <- "输出_1号梯LEDf"
   Rectangle "矩形_197" at 427,186 size 18x4
      Appearance <- "输出_1号梯LEDa"
   Rectangle "矩形_198" at 424,190 size 4x18
      Appearance <- "输出_1号梯LEDe"
   Rectangle "矩形_199" at 427,208 size 18x4
      Appearance <- "输出_1号梯LEDd"
   Rectangle "矩形_200" at 444,168 size 4x18
      Appearance <- "输出_1号梯LEDb"
   Rectangle "矩形_201" at 444,190 size 4x18
      Appearance <- "输出_1号梯LEDc"
   Rectangle "矩形_35" at 555,170 size 4x18
      Appearance <- "输出_2号梯LEDi"
   Rectangle "矩形_36" at 555,192 size 4x18
      Appearance <- "输出_2号梯LEDj"
   Rectangle "矩形_37" at 568,168 size 18x4
      Appearance <- "输出_2号梯LEDa"
   Rectangle "矩形_38" at 565,172 size 4x18
      Appearance <- "输出_2号梯LEDf"
   Rectangle "矩形_39" at 568,189 size 18x4
      Appearance <- "输出_2号梯LEDg"
   Rectangle "矩形_40" at 565,193 size 4x18
      Appearance <- "输出_2号梯LEDe"
   Rectangle "矩形_41" at 568,211 size 18x4
      Appearance <- "输出_2号梯LEDd"
   Rectangle "矩形_42" at 585,171 size 4x18
      Appearance <- "输出_2号梯LEDb"
   Rectangle "矩形_43" at 585,193 size 4x18
      Appearance <- "输出_2号梯LEDc"
   Rectangle "矩形_7" at 416,295 size 4x18
      Appearance <- "输出_3号梯LEDi"
   Rectangle "矩形_8" at 416,317 size 4x18
      Appearance <- "输出_3号梯LEDj"
   Rectangle "矩形_9" at 429,293 size 18x4
      Appearance <- "输出_3号梯LEDa"
   Rectangle "矩形_10" at 426,297 size 4x18
      Appearance <- "输出_3号梯LEDf"
   Rectangle "矩形_11" at 429,314 size 18x4
      Appearance <- "输出_3号梯LEDg"
   Rectangle "矩形_12" at 426,318 size 4x18
      Appearance <- "输出_3号梯LEDe"
   Rectangle "矩形_13" at 429,336 size 18x4
      Appearance <- "输出_3号梯LEDd"
   Rectangle "矩形_14" at 446,296 size 4x18
      Appearance <- "输出_3号梯LEDb"
   Rectangle "矩形_15" at 446,318 size 4x18
      Appearance <- "输出_3号梯LEDc"
   Rectangle "矩形_49" at 556,299 size 4x18
      Appearance <- "输出_4号梯LEDi"
   Rectangle "矩形_50" at 556,321 size 4x18
      Appearance <- "输出_4号梯LEDj"
   Rectangle "矩形_51" at 569,297 size 18x4
      Appearance <- "输出_4号梯LEDa"
   Rectangle "矩形_52" at 566,301 size 4x18
      Appearance <- "输出_4号梯LEDf"
   Rectangle "矩形_53" at 569,318 size 18x4
      Appearance <- "输出_4号梯LEDg"
   Rectangle "矩形_54" at 566,322 size 4x18
      Appearance <- "输出_4号梯LEDe"
   Rectangle "矩形_55" at 569,340 size 18x4
      Appearance <- "输出_4号梯LEDd"
   Rectangle "矩形_56" at 586,300 size 4x18
      Appearance <- "输出_4号梯LEDb"
   Rectangle "矩形_57" at 586,322 size 4x18
      Appearance <- "输出_4号梯LEDc"
   Rectangle "矩形_21" at 419,437 size 4x18
      Appearance <- "输出_5号梯LEDi"
   Rectangle "矩形_22" at 419,459 size 4x18
      Appearance <- "输出_5号梯LEDj"
   Rectangle "矩形_23" at 432,435 size 18x4
      Appearance <- "输出_5号梯LEDa"
   Rectangle "矩形_24" at 429,439 size 4x18
      Appearance <- "输出_5号梯LEDf"
   Rectangle "矩形_25" at 432,456 size 18x4
      Appearance <- "输出_5号梯LEDg"
   Rectangle "矩形_26" at 429,460 size 4x18
      Appearance <- "输出_5号梯LEDe"
   Rectangle "矩形_27" at 432,478 size 18x4
      Appearance <- "输出_5号梯LEDd"
   Rectangle "矩形_28" at 449,438 size 4x18
      Appearance <- "输出_5号梯LEDb"
   Rectangle "矩形_29" at 449,460 size 4x18
      Appearance <- "输出_5号梯LEDc"
   Rectangle "矩形_63" at 558,436 size 4x18
      Appearance <- "输出_6号梯LEDi"
   Rectangle "矩形_64" at 558,458 size 4x18
      Appearance <- "输出_6号梯LEDj"
   Rectangle "矩形_65" at 571,434 size 18x4
      Appearance <- "输出_6号梯LEDa"
   Rectangle "矩形_66" at 568,438 size 4x18
      Appearance <- "输出_6号梯LEDf"
   Rectangle "矩形_67" at 571,455 size 18x4
      Appearance <- "输出_6号梯LEDg"
   Rectangle "矩形_68" at 568,459 size 4x18
      Appearance <- "输出_6号梯LEDe"
   Rectangle "矩形_69" at 571,477 size 18x4
      Appearance <- "输出_6号梯LEDd"
   Rectangle "矩形_70" at 588,437 size 4x18
      Appearance <- "输出_6号梯LEDb"
   Rectangle "矩形_71" at 588,459 size 4x18
      Appearance <- "输出_6号梯LEDc"
   Polygon "多边形_5" at 335,169 size 32x16
      Appearance <- "输出_1号梯下行指示"
   Polygon "多边形_6" at 335,188 size 32x16
      Appearance <- "输出_1号梯上行指示"
   Polygon "多边形_1" at 337,298 size 32x16
      Appearance <- "输出_3号梯下行指示"
   Polygon "多边形_2" at 337,317 size 32x16
      Appearance <- "输出_3号梯上行指示"
   Polygon "多边形_3" at 335,435 size 32x16
      Appearance <- "输出_5号梯下行指示"
   Polygon "多边形_4" at 335,454 size 32x16
      Appearance <- "输出_5号梯上行指示"
   Polygon "多边形_7" at 484,440 size 32x16
      Appearance <- "输出_6号梯下行指示"
   Polygon "多边形_8" at 484,459 size 32x16
      Appearance <- "输出_6号梯上行指示"
   Polygon "多边形_9" at 484,305 size 32x16
      Appearance <- "输出_4号梯下行指示"
   Polygon "多边形_10" at 484,324 size 32x16
      Appearance <- "输出_4号梯上行指示"
   Polygon "多边形_11" at 484,170 size 32x16
      Appearance <- "输出_2号梯下行指示"
   Polygon "多边形_12" at 484,189 size 32x16
      Appearance <- "输出_2号梯上行指示"
   Polygon "多边形_13" at 123,83 size 32x16
      Appearance <- "输出_10层下行呼梯按钮指示灯"
   Polygon "多边形_14" at 123,513 size 32x16
      Appearance <- "输出_1层上行呼梯按钮指示灯"
   Polygon "多边形_15" at 155,473 size 32x16
      Appearance <- "输出_2层下行呼梯按钮指示灯"
   Polygon "多边形_16" at 91,469 size 32x16
      Appearance <- "输出_2层上行呼梯按钮指示灯"
   Polygon "多边形_17" at 155,423 size 32x16
      Appearance <- "输出_3层下行呼梯按钮指示灯"
   Polygon "多边形_18" at 91,419 size 32x16
      Appearance <- "输出_3层上行呼梯按钮指示灯"
   Polygon "多边形_19" at 155,373 size 32x16
      Appearance <- "输出_4层下行呼梯按钮指示灯"
   Polygon "多边形_20" at 91,369 size 32x16
      Appearance <- "输出_4层上行呼梯按钮指示灯"
   Polygon "多边形_21" at 155,323 size 32x16
      Appearance <- "输出_5层下行呼梯按钮指示灯"
   Polygon "多边形_22" at 91,319 size 32x16
      Appearance <- "输出_5层上行呼梯按钮指示灯"
   Polygon "多边形_23" at 155,273 size 32x16
      Appearance <- "输出_6层下行呼梯按钮指示灯"
   Polygon "多边形_24" at 91,269 size 32x16
      Appearance <- "输出_6层上行呼梯按钮指示灯"
   Polygon "多边形_25" at 155,223 size 32x16
      Appearance <- "输出_7层下行呼梯按钮指示灯"
   Polygon "多边形_26" at 91,219 size 32x16
      Appearance <- "输出_7层上行呼梯按钮指示灯"
   Polygon "多边形_27" at 155,173 size 32x16
      Appearance <- "输出_8层下行呼梯按钮指示灯"
   Polygon "多边形_28" at 91,169 size 32x16
      Appearance <- "输出_8层上行呼梯按钮指示灯"
   Polygon "多边形_29" at 155,123 size 32x16
      Appearance <- "输出_9层下行呼梯按钮指示灯"
   Polygon "多边形_30" at 91,119 size 32x16
      Appearance <- "输出_9层上行呼梯按钮指示灯"
   Clock "时钟_1" at 664,57 size 101x57
   DateTimeField "日期/时间域_1" at 491,71 size 184x28

screen "用户设置" 800x600
   Button "按钮_7" at 554,513 size 110x66; TextOff '主画面'
      on Click: ActivateScreen("主画面", 0)
   TextField "文本域_1" at 385,17 size 210x27; Text '-- 用户设置'
   TextField "文本域_3" at 85,12 size 292x31; Text '电 梯 监 控 系 统'
   Button "按钮_1" at 674,513 size 106x66; TextOff '退出系统'
      on Click: StopRuntime(0)
   UserView "用户视图_1" at 116,172 size 558x230
   Clock "时钟_1" at 664,57 size 101x57
   DateTimeField "日期/时间域_1" at 491,71 size 184x28

screen "电梯状态总览画面" 800x600
   Button "按钮_7" at 555,518 size 110x66; TextOff '主画面'
      on Click: ActivateScreen("主画面", 0)
   Button "按钮_8" at 672,517 size 106x67; TextOff '退出系统'
      on Click: StopRuntime(0)
   TextField "文本域_1" at 440,13 size 263x31; Text '--电梯状态总览'
   Button "按钮_1" at 176,142 size 202x49; TextOff '#1电梯'
      on Click: ActivateScreen("1#电梯状态画面", 0)
   Button "按钮_2" at 412,216 size 202x49; TextOff '#4电梯'
      on Click: ActivateScreen("4#电梯状态画面", 0)
   Button "按钮_3" at 411,144 size 202x49; TextOff '#2电梯'
      on Click: ActivateScreen("2#电梯状态画面", 0)
   Button "按钮_4" at 177,216 size 202x49; TextOff '#3电梯'
      on Click: ActivateScreen("3#电梯状态画面", 0)
   Button "按钮_5" at 179,286 size 202x49; TextOff '#5电梯'
      on Click: ActivateScreen("5#电梯状态画面", 0)
   Button "按钮_6" at 412,286 size 202x49; TextOff '#6电梯'
      on Click: ActivateScreen("6#电梯状态画面", 0)
   TextField "文本域_3" at 141,12 size 323x31; Text '电 梯 监 控 系 统'
   Clock "时钟_1" at 664,57 size 101x57
   DateTimeField "日期/时间域_1" at 491,71 size 184x28

screen "电梯运行监控画面1" 800x600
   Button "按钮_2" at 72,133 size 88x45; TextOff 'Text'
      on Click: ActivateScreen("电梯运行监控画面1", 0)
   Button "按钮_7" at 559,517 size 110x68; TextOff '主画面'
      on Click: ActivateScreen("主画面", 0)
   TextField "文本域_1" at 385,17 size 274x27; Text '-- 1#电梯运行监控'
   TextField "文本域_3" at 81,12 size 296x31; Text '电 梯 监 控 系 统'
   Button "按钮_1" at 678,516 size 106x68; TextOff '退出系统'
      on Click: StopRuntime(0)
   Circle "圆_1" at 21,138 size 35x35
      Appearance <- "1号梯正常运行"
   TextField "文本域_2" at 85,141 size 68x29; Text '1#电梯'
   Circle "圆_7" at 199,171 size 31x31
      Appearance <- "输出_1号梯1层按钮指示灯"
   TextField "文本域_9" at 208,175 size 14x19; Text '1'
   Circle "圆_8" at 247,171 size 31x31
      Appearance <- "输出_1号梯2层按钮指示灯"
   TextField "文本域_10" at 256,175 size 14x19; Text '2'
   Circle "圆_9" at 295,171 size 31x31
      Appearance <- "输出_1号梯3层按钮指示灯"
   TextField "文本域_11" at 304,175 size 14x19; Text '3'
   Circle "圆_10" at 199,221 size 31x31
      Appearance <- "输出_1号梯4层按钮指示灯"
   TextField "文本域_12" at 208,225 size 14x19; Text '4'
   Circle "圆_11" at 247,221 size 31x31
      Appearance <- "输出_1号梯5层按钮指示灯"
   TextField "文本域_13" at 256,225 size 14x19; Text '5'
   Circle "圆_12" at 295,221 size 31x31
      Appearance <- "输出_1号梯6层按钮指示灯"
   TextField "文本域_14" at 304,225 size 14x19; Text '6'
   Circle "圆_13" at 199,271 size 31x31
      Appearance <- "输出_1号梯7层按钮指示灯"
   TextField "文本域_15" at 208,275 size 14x19; Text '7'
   Circle "圆_14" at 247,271 size 31x31
      Appearance <- "输出_1号梯8层按钮指示灯"
   TextField "文本域_16" at 256,275 size 14x19; Text '8'
   Circle "圆_15" at 295,271 size 31x31
      Appearance <- "输出_1号梯9层按钮指示灯"
   TextField "文本域_17" at 304,275 size 14x19; Text '9'
   Circle "圆_16" at 248,317 size 31x31
      Appearance <- "输出_1号梯10层按钮指示灯"
   TextField "文本域_18" at 252,322 size 23x19; Text '10'
   TextField "文本域_19" at 368,345 size 61x19; Text '开门'
   TextField "文本域_20" at 457,347 size 53x19; Text '关门'
   TextField "文本域_21" at 528,284 size 95x25; Text '运行方向：'
   TextField "文本域_22" at 529,348 size 94x24; Text '厢门状态：'
   Rectangle "矩形_2" at 178,400 size 599x88
      Visibility <- "输入_1号梯检修信号"
   GraphicView "图形视图_1" at 609,139 size 124x108; Picture "b_95950E8D4E6480C12C2CE472E64CCEF4[1]"
   Polygon "多边形_3" at 372,298 size 16x33
      Appearance <- "输出_1号梯开门继电器"
   Polygon "多边形_4" at 392,298 size 16x33
      Appearance <- "输出_1号梯开门继电器"
   Polygon "多边形_7" at 459,298 size 16x32
      Appearance <- "输出_1号梯关门继电器"
   Polygon "多边形_8" at 479,298 size 16x32
      Appearance <- "输出_1号梯关门继电器"
   TextField "文本域_24" at 620,299 size 44x19; Text '上行'
      Visibility <- "输出_1号梯上行指示"
   TextField "文本域_25" at 678,297 size 44x19; Text '下行'
      Visibility <- "输出_1号梯下行指示"
   TextField "文本域_27" at 641,361 size 52x19; Text '开启'
      Visibility <- "输出_1号梯开门继电器"
   TextField "文本域_28" at 706,361 size 52x19; Text '关闭'
      Visibility <- "输出_1号梯关门继电器"
   Button "按钮_3" at 72,189 size 88x45; TextOff 'Text'
      on Click: ActivateScreen("电梯运行监控画面2", 0)
   Circle "圆_2" at 21,194 size 35x35
      Appearance <- "2号梯正常运行"
   TextField "文本域_4" at 84,194 size 68x29; Text '2#电梯'
   Button "按钮_4" at 72,247 size 88x45; TextOff 'Text'
      on Click: ActivateScreen("电梯运行监控画面3", 0)
   Circle "圆_3" at 21,252 size 35x35
      Appearance <- "3号梯正常运行"
   TextField "文本域_5" at 85,252 size 68x29; Text '3#电梯'
   Button "按钮_5" at 72,305 size 88x45; TextOff 'Text'
      on Click: ActivateScreen("电梯运行监控画面4", 0)
   Circle "圆_4" at 21,310 size 35x35
      Appearance <- "4号梯正常运行"
   TextField "文本域_6" at 84,310 size 68x29; Text '4#电梯'
   Button "按钮_6" at 72,363 size 88x45; TextOff 'Text'
      on Click: ActivateScreen("电梯运行监控画面5", 0)
   Circle "圆_5" at 21,368 size 35x35
      Appearance <- "5号梯正常运行"
   TextField "文本域_7" at 80,371 size 68x29; Text '5#电梯'
   Button "按钮_8" at 72,421 size 88x45; TextOff 'Text'
      on Click: ActivateScreen("电梯运行监控画面6", 0)
   Circle "圆_6" at 21,426 size 35x35
      Appearance <- "6号梯正常运行"
   TextField "文本域_8" at 82,427 size 68x29; Text '6#电梯'
   Rectangle "矩形_193" at 521,167 size 4x18
      Appearance <- "输出_1号梯LEDi"
   Rectangle "矩形_194" at 521,189 size 4x18
      Appearance <- "输出_1号梯LEDj"
   Rectangle "矩形_195" at 534,165 size 18x4
      Appearance <- "输出_1号梯LEDa"
   Rectangle "矩形_196" at 531,169 size 4x18
      Appearance <- "输出_1号梯LEDf"
   Rectangle "矩形_197" at 534,186 size 18x4
      Appearance <- "输出_1号梯LEDg"
   Rectangle "矩形_198" at 531,190 size 4x18
      Appearance <- "输出_1号梯LEDe"
   Rectangle "矩形_199" at 534,208 size 18x4
      Appearance <- "输出_1号梯LEDd"
   Rectangle "矩形_200" at 551,168 size 4x18
      Appearance <- "输出_1号梯LEDb"
   Rectangle "矩形_201" at 551,190 size 4x18
      Appearance <- "输出_1号梯LEDc"
   Rectangle "矩形_3" at 426,152 size 6x34
      Appearance <- "输出_1号梯上行指示"
   Polygon "多边形_5" at 414,148 size 15x17
      Appearance <- "输出_1号梯上行指示"
   Polygon "多边形_6" at 429,148 size 14x17
      Appearance <- "输出_1号梯上行指示"
   Rectangle "矩形_73" at 426,187 size 6x34
      Appearance <- "输出_1号梯下行指示"
   Polygon "多边形_1" at 412,209 size 17x15
      Appearance <- "输出_1号梯下行指示"
   Polygon "多边形_2" at 429,209 size 17x15
      Appearance <- "输出_1号梯下行指示"
   TextField "文本域_23" at 343,413 size 309x70; Text '1#正常运行'
      Visibility <- "1号梯正常运行"
   TextField "文本域_32" at 346,414 size 309x70; Text '1#满载故障'
      Visibility <- "输出_1号梯满载指示"
   TextField "文本域_33" at 343,410 size 309x74; Text '1#检修故障'
      Visibility <- "输入_1号梯检修信号"
   Polygon "多边形_28" at 620,276 size 32x16
      Visibility <- "输出_1号梯上行指示"
   Polygon "多边形_27" at 681,276 size 32x16
      Visibility <- "输出_1号梯下行指示"
   Circle "圆_18" at 650,338 size 21x21
      Visibility <- "输出_1号梯开门继电器"
   Circle "圆_19" at 714,338 size 21x21
      Visibility <- "输出_1号梯关门继电器"
   Clock "时钟_1" at 665,53 size 101x57
   DateTimeField "日期/时间域_1" at 491,71 size 184x28
   IOField "I/O 域_1" at 110,507 size 96x32; FormatPattern s99999
      ProcessValue <- "1号梯载重量"
   TextField "文本域_26" at 23,498 size 84x47; Text '当前重量'

screen "电梯运行监控画面2" 800x600
   Button "按钮_7" at 559,517 size 110x68; TextOff '主画面'
      on Click: ActivateScreen("主画面", 0)
   TextField "文本域_1" at 385,17 size 285x27; Text '-- 2#电梯运行监控'
   TextField "文本域_3" at 114,12 size 263x31; Text '电 梯 监 控 系 统'
   Button "按钮_1" at 678,516 size 106x68; TextOff '退出系统'
      on Click: StopRuntime(0)
   Circle "圆_7" at 199,171 size 31x31
      Appearance <- "输出_2号梯1层按钮指示灯"
   TextField "文本域_9" at 208,175 size 14x19; Text '1'
   Circle "圆_8" at 247,171 size 31x31
      Appearance <- "输出_2号梯2层按钮指示灯"
   TextField "文本域_10" at 256,175 size 14x19; Text '2'
   Circle "圆_9" at 295,171 size 31x31
      Appearance <- "输出_2号梯3层按钮指示灯"
   TextField "文本域_11" at 304,175 size 14x19; Text '3'
   Circle "圆_10" at 199,221 size 31x31
      Appearance <- "输出_2号梯4层按钮指示灯"
   TextField "文本域_12" at 208,225 size 14x19; Text '4'
   Circle "圆_11" at 247,221 size 31x31
      Appearance <- "输出_2号梯5层按钮指示灯"
   TextField "文本域_13" at 256,225 size 14x19; Text '5'
   Circle "圆_12" at 295,221 size 31x31
      Appearance <- "输出_2号梯6层按钮指示灯"
   TextField "文本域_14" at 304,225 size 14x19; Text '6'
   Circle "圆_13" at 199,271 size 31x31
      Appearance <- "输出_2号梯7层按钮指示灯"
   TextField "文本域_15" at 208,275 size 14x19; Text '7'
   Circle "圆_14" at 247,271 size 31x31
      Appearance <- "输出_2号梯8层按钮指示灯"
   TextField "文本域_16" at 256,275 size 14x19; Text '8'
   Circle "圆_15" at 295,271 size 31x31
      Appearance <- "输出_2号梯9层按钮指示灯"
   TextField "文本域_17" at 304,275 size 14x19; Text '9'
   Circle "圆_16" at 248,317 size 31x31
      Appearance <- "输出_2号梯10层按钮指示灯"
   TextField "文本域_18" at 252,322 size 23x19; Text '10'
   TextField "文本域_19" at 368,345 size 61x19; Text '开门'
   TextField "文本域_20" at 457,347 size 53x19; Text '关门'
   TextField "文本域_21" at 528,289 size 95x25; Text '运行方向：'
   TextField "文本域_22" at 529,349 size 94x24; Text '厢门状态：'
   TextField "文本域_23" at 343,408 size 309x70; Text '2#正常运行'
      Visibility <- "2号梯正常运行"
   GraphicView "图形视图_1" at 609,139 size 124x108; Picture "b_95950E8D4E6480C12C2CE472E64CCEF4[1]"
   Polygon "多边形_3" at 372,298 size 16x33
      Appearance <- "输出_2号梯开门继电器"
   Polygon "多边形_4" at 392,298 size 16x33
      Appearance <- "输出_2号梯开门继电器"
   Polygon "多边形_7" at 459,298 size 16x32
      Appearance <- "输出_2号梯关门继电器"
   Polygon "多边形_8" at 479,298 size 16x32
      Appearance <- "输出_2号梯关门继电器"
   TextField "文本域_24" at 620,301 size 44x19; Text '上行'
      Visibility <- "输出_1号梯上行指示"
   TextField "文本域_25" at 675,300 size 44x19; Text '下行'
      Visibility <- "输出_1号梯下行指示"
   TextField "文本域_27" at 641,355 size 52x19; Text '开启'
      Visibility <- "输出_2号梯开门继电器"
   TextField "文本域_28" at 705,356 size 52x19; Text '关闭'
      Visibility <- "输出_2号梯关门继电器"
   Polygon "多边形_28" at 620,279 size 32x16
      Visibility <- "输出_1号梯上行指示"
   Polygon "多边形_27" at 678,279 size 32x16
      Visibility <- "输出_1号梯下行指示"
   Circle "圆_18" at 650,334 size 21x21
      Visibility <- "输出_2号梯开门继电器"
   Circle "圆_19" at 713,335 size 21x21
      Visibility <- "输出_2号梯关门继电器"
   Button "按钮_2" at 72,133 size 88x45; TextOff 'Text'
      on Click: ActivateScreen("电梯运行监控画面1", 0)
   TextField "文本域_2" at 84,131 size 68x29; Text '1#电梯'
   Button "按钮_3" at 72,189 size 88x45; TextOff 'Text'
      on Click: ActivateScreen("电梯运行监控画面2", 0)
   TextField "文本域_4" at 84,187 size 68x29; Text '2#电梯'
   Button "按钮_4" at 72,247 size 88x45; TextOff 'Text'
      on Click: ActivateScreen("电梯运行监控画面3", 0)
   TextField "文本域_5" at 84,245 size 68x29; Text '3#电梯'
   Button "按钮_5" at 72,305 size 88x45; TextOff 'Text'
      on Click: ActivateScreen("电梯运行监控画面4", 0)
   TextField "文本域_6" at 84,303 size 68x29; Text '4#电梯'
   Button "按钮_6" at 72,363 size 88x45; TextOff 'Text'
      on Click: ActivateScreen("电梯运行监控画面5", 0)
   TextField "文本域_7" at 84,361 size 68x29; Text '5#电梯'
   Button "按钮_8" at 72,421 size 88x45; TextOff 'Text'
      on Click: ActivateScreen("电梯运行监控画面6", 0)
   TextField "文本域_8" at 84,419 size 68x29; Text '6#电梯'
   Rectangle "矩形_193" at 524,163 size 4x18
      Appearance <- "输出_2号梯LEDi"
   Rectangle "矩形_194" at 524,185 size 4x18
      Appearance <- "输出_2号梯LEDj"
   Rectangle "矩形_195" at 537,161 size 18x4
      Appearance <- "输出_2号梯LEDa"
   Rectangle "矩形_196" at 534,165 size 4x18
      Appearance <- "输出_2号梯LEDf"
   Rectangle "矩形_197" at 537,182 size 18x4
      Appearance <- "输出_2号梯LEDg"
   Rectangle "矩形_198" at 534,186 size 4x18
      Appearance <- "输出_2号梯LEDe"
   Rectangle "矩形_199" at 537,204 size 18x4
      Appearance <- "输出_2号梯LEDd"
   Rectangle "矩形_200" at 554,164 size 4x18
      Appearance <- "输出_2号梯LEDb"
   Rectangle "矩形_201" at 554,186 size 4x18
      Appearance <- "输出_2号梯LEDc"
   Rectangle "矩形_72" at 429,147 size 6x34
      Appearance <- "输出_2号梯上行指示"
   Polygon "多边形_5" at 417,143 size 15x17
      Appearance <- "输出_2号梯上行指示"
   Polygon "多边形_6" at 432,143 size 14x17
      Appearance <- "输出_2号梯上行指示"
   Rectangle "矩形_73" at 429,182 size 6x34
      Appearance <- "输出_2号梯下行指示"
   Polygon "多边形_1" at 415,204 size 17x15
      Appearance <- "输出_2号梯下行指示"
   Polygon "多边形_2" at 432,204 size 17x15
      Appearance <- "输出_2号梯下行指示"
   Circle "圆_1" at 21,138 size 35x35
      Appearance <- "1号梯正常运行"
   Circle "圆_2" at 21,194 size 35x35
      Appearance <- "2号梯正常运行"
   Circle "圆_3" at 21,252 size 35x35
      Appearance <- "3号梯正常运行"
   Circle "圆_4" at 21,310 size 35x35
      Appearance <- "4号梯正常运行"
   Circle "圆_5" at 21,368 size 35x35
      Appearance <- "5号梯正常运行"
   Circle "圆_6" at 21,426 size 35x35
      Appearance <- "6号梯正常运行"
   TextField "文本域_33" at 343,410 size 309x70; Text '2#检修故障'
      Visibility <- "输入_2号梯检修信号"
   TextField "文本域_32" at 345,410 size 309x70; Text '2#满载故障'
      Visibility <- "输出_2号梯满载指示"
   Clock "时钟_1" at 664,57 size 101x57
   DateTimeField "日期/时间域_1" at 491,71 size 184x28
   TextField "文本域_26" at 23,498 size 84x47; Text '当前重量'
   IOField "I/O 域_1" at 110,507 size 96x32; FormatPattern s99999
      ProcessValue <- "2号梯载重量"

screen "电梯运行监控画面3" 800x600
   Button "按钮_7" at 559,517 size 110x68; TextOff '主画面'
      on Click: ActivateScreen("主画面", 0)
   TextField "文本域_1" at 385,17 size 304x27; Text '-- 3#电梯运行监控'
   TextField "文本域_3" at 114,12 size 263x31; Text '电 梯 监 控 系 统'
   Button "按钮_1" at 678,516 size 106x68; TextOff '退出系统'
      on Click: StopRuntime(0)
   Circle "圆_7" at 199,171 size 31x31
      Appearance <- "输出_3号梯1层按钮指示灯"
   TextField "文本域_9" at 208,175 size 14x19; Text '1'
   Circle "圆_8" at 247,171 size 31x31
      Appearance <- "输出_3号梯2层按钮指示灯"
   TextField "文本域_10" at 256,175 size 14x19; Text '2'
   Circle "圆_9" at 295,171 size 31x31
      Appearance <- "输出_3号梯3层按钮指示灯"
   TextField "文本域_11" at 304,175 size 14x19; Text '3'
   Circle "圆_10" at 199,221 size 31x31
      Appearance <- "输出_3号梯4层按钮指示灯"
   TextField "文本域_12" at 208,225 size 14x19; Text '4'
   Circle "圆_11" at 247,221 size 31x31
      Appearance <- "输出_3号梯5层按钮指示灯"
   TextField "文本域_13" at 256,225 size 14x19; Text '5'
   Circle "圆_12" at 295,221 size 31x31
      Appearance <- "输出_3号梯6层按钮指示灯"
   TextField "文本域_14" at 304,225 size 14x19; Text '6'
   Circle "圆_13" at 199,271 size 31x31
      Appearance <- "输出_3号梯7层按钮指示灯"
   TextField "文本域_15" at 208,275 size 14x19; Text '7'
   Circle "圆_14" at 247,271 size 31x31
      Appearance <- "输出_3号梯8层按钮指示灯"
   TextField "文本域_16" at 256,275 size 14x19; Text '8'
   Circle "圆_15" at 295,271 size 31x31
      Appearance <- "输出_3号梯9层按钮指示灯"
   TextField "文本域_17" at 304,275 size 14x19; Text '9'
   Circle "圆_16" at 248,317 size 31x31
      Appearance <- "输出_3号梯10层按钮指示灯"
   TextField "文本域_18" at 252,322 size 23x19; Text '10'
   TextField "文本域_19" at 368,345 size 61x19; Text '开门'
   TextField "文本域_20" at 457,347 size 53x19; Text '关门'
   TextField "文本域_21" at 528,277 size 95x25; Text '运行方向：'
   TextField "文本域_22" at 529,337 size 94x24; Text '厢门状态：'
   TextField "文本域_23" at 341,406 size 309x70; Text '3#正常运行'
      Visibility <- "3号梯正常运行"
   GraphicView "图形视图_1" at 609,139 size 124x108; Picture "b_95950E8D4E6480C12C2CE472E64CCEF4[1]"
   Polygon "多边形_3" at 372,298 size 16x33
      Appearance <- "输出_3号梯开门继电器"
   Polygon "多边形_4" at 392,298 size 16x33
      Appearance <- "输出_3号梯开门继电器"
   Polygon "多边形_7" at 459,298 size 16x32
      Appearance <- "输出_3号梯关门继电器"
   Polygon "多边形_8" at 479,298 size 16x32
      Appearance <- "输出_3号梯关门继电器"
   TextField "文本域_24" at 620,287 size 44x19; Text '上行'
      Visibility <- "输出_3号梯上行指示"
   TextField "文本域_25" at 676,285 size 44x19; Text '下行'
      Visibility <- "输出_3号梯下行指示"
   TextField "文本域_27" at 641,346 size 52x19; Text '开启'
      Visibility <- "输出_3号梯开门继电器"
   TextField "文本域_28" at 705,345 size 52x19; Text '关闭'
      Visibility <- "输出_3号梯关门继电器"
   Polygon "多边形_28" at 620,264 size 32x16
      Visibility <- "输出_3号梯上行指示"
   Polygon "多边形_27" at 679,264 size 32x16
      Visibility <- "输出_3号梯下行指示"
   Circle "圆_18" at 649,325 size 21x21
      Visibility <- "输出_3号梯开门继电器"
   Circle "圆_19" at 712,324 size 21x21
      Visibility <- "输出_3号梯关门继电器"
   Button "按钮_2" at 72,133 size 88x45; TextOff 'Text'
      on Click: ActivateScreen("电梯运行监控画面1", 0)
   TextField "文本域_2" at 84,137 size 68x29; Text '1#电梯'
   Button "按钮_3" at 72,189 size 88x45; TextOff 'Text'
      on Click: ActivateScreen("电梯运行监控画面2", 0)
   TextField "文本域_4" at 84,196 size 68x29; Text '2#电梯'
   Button "按钮_4" at 72,247 size 88x45; TextOff 'Text'
      on Click: ActivateScreen("电梯运行监控画面3", 0)
   TextField "文本域_5" at 81,256 size 68x29; Text '3#电梯'
   Button "按钮_5" at 72,305 size 88x45; TextOff 'Text'
      on Click: ActivateScreen("电梯运行监控画面4", 0)
   TextField "文本域_6" at 81,310 size 68x29; Text '4#电梯'
   Button "按钮_6" at 72,363 size 88x45; TextOff 'Text'
      on Click: ActivateScreen("电梯运行监控画面5", 0)
   TextField "文本域_7" at 81,368 size 68x29; Text '5#电梯'
   Button "按钮_8" at 72,421 size 88x45; TextOff 'Text'
      on Click: ActivateScreen("电梯运行监控画面6", 0)
   TextField "文本域_8" at 81,426 size 68x29; Text '6#电梯'
   Rectangle "矩形_193" at 528,160 size 4x18
      Appearance <- "输出_3号梯LEDi"
   Rectangle "矩形_194" at 528,182 size 4x18
      Appearance <- "输出_3号梯LEDj"
   Rectangle "矩形_195" at 541,158 size 18x4
      Appearance <- "输出_3号梯LEDa"
   Rectangle "矩形_196" at 538,162 size 4x18
      Appearance <- "输出_3号梯LEDf"
   Rectangle "矩形_197" at 541,179 size 18x4
      Appearance <- "输出_3号梯LEDg"
   Rectangle "矩形_198" at 538,183 size 4x18
      Appearance <- "输出_3号梯LEDe"
   Rectangle "矩形_199" at 541,201 size 18x4
      Appearance <- "输出_3号梯LEDd"
   Rectangle "矩形_200" at 558,161 size 4x18
      Appearance <- "输出_3号梯LEDb"
   Rectangle "矩形_201" at 558,183 size 4x18
      Appearance <- "输出_3号梯LEDc"
   Rectangle "矩形_72" at 431,153 size 6x34
      Appearance <- "输出_3号梯上行指示"
   Polygon "多边形_5" at 419,149 size 15x17
      Appearance <- "输出_3号梯上行指示"
   Polygon "多边形_6" at 434,149 size 14x17
      Appearance <- "输出_3号梯上行指示"
   Rectangle "矩形_73" at 431,188 size 6x34
      Appearance <- "输出_3号梯下行指示"
   Polygon "多边形_1" at 417,210 size 17x15
      Appearance <- "输出_3号梯下行指示"
   Polygon "多边形_2" at 434,210 size 17x15
      Appearance <- "输出_3号梯下行指示"
   Circle "圆_1" at 21,138 size 35x35
      Appearance <- "1号梯正常运行"
   Circle "圆_2" at 21,194 size 35x35
      Appearance <- "2号梯正常运行"
   Circle "圆_3" at 21,252 size 35x35
      Appearance <- "3号梯正常运行"
   Circle "圆_4" at 21,310 size 35x35
      Appearance <- "4号梯正常运行"
   Circle "圆_5" at 21,368 size 35x35
      Appearance <- "5号梯正常运行"
   Circle "圆_6" at 21,426 size 35x35
      Appearance <- "6号梯正常运行"
   TextField "文本域_33" at 343,406 size 309x70; Text '3#检修故障'
      Visibility <- "输入_3号梯检修信号"
   TextField "文本域_32" at 340,408 size 309x70; Text '3#满载故障'
      Visibility <- "输出_3号梯满载指示"
   Clock "时钟_1" at 664,57 size 101x57
   DateTimeField "日期/时间域_1" at 491,71 size 184x28
   TextField "文本域_26" at 23,498 size 84x47; Text '当前重量'
   IOField "I/O 域_1" at 110,507 size 96x32; FormatPattern s99999
      ProcessValue <- "3号梯载重量"

